(* IEC 61131-3 sources: daoli-st-library/DL_Process (part 37) *)

(* ---- FB_DL_HjtPvdSeq.st ---- *)
(*
  FB_DL_HjtPvdSeq  —  HJT 光伏 PVD 镀膜腔体顺控 / HJT PVD coating chamber sequence
  分类 Category : DL_Process
  码位 Code     : 16#06_0_B6
  段位说明      : R38 W7 预留 B6~BF 本轮正式启用，本件启用 B6 格
  版本 Version  : 1.0.0
  来源 Source   : 自研线（半导体/光伏工艺）— HJT PVD 镀膜公开工艺段序
  溯源 Origin   : clean-room 实现，未复制任何源码行
                  （段序语义对齐 FB_DL_StepSequencer，不实例化；接口契约按 I_DL_* 真实成员名调用）
  功能 Function : 1) 四段顺控 BaseVac→Preheat→Coat→Unload，段尾经 Done 回 Idle；
                  2) 本底真空段：抽气至 fBaseVacKpa（深度判据）；
                  3) 预热段：温区 SetSetpoint 到位 + 配方时长驻留；
                  4) 工艺镀膜段：真空深度与温度双到位联锁内置（联锁不满足只等待不故障），
                  配方时长到点收段；
                  5) 取片段：放气常压确认 AND bUnloadPermit 联锁双确认才进 Done；
                  6) 段超时升级：四段各配独立超时 TON，超时锁故障。
  边界 Boundary : ① 真空接口契约：iVac.fPressure 为负压值，深度 = −fPressure（取正深度比较）；
                  ② 组态域闸覆盖全部参与换算引脚（R151）；配方/超时全 0 判组态错；
                  ③ R228-A 达标声明：八只 TON 均单相独占（IN 为单相等式），跨相迁移拍 IN 必断；
                  ④ R228-B 达标声明：eFault 迁出 = rtReset.Q（输入引脚，恒可达），逐字写于此；
                  ⑤ 解除式自证：段超时故障解除 = bReset 上升沿 AND eState = Idle（迁出边唯一可达）；
                  ⑥ CASE 全态覆盖 + ELSE 兜底置 Fault。
  依赖 Depends  : I_DL_VacuumGenerator / I_DL_TemperatureZone（注入，不实例化）；
                  段序语义对齐 FB_DL_StepSequencer（已注册，不实例化）
  码表 Error codes（本件格 06_0_B6，子码步进 +0x100）:
    16#0006_01B6 信息级：周期完成（Done 相）
    16#0006_02B6 故障级：组态非法（真空目标/温度目标/容差/常压阈/配方/超时域非法），锁存至复位
    16#0006_03B6 故障级：段超时升级（四段独立计时），锁存至复位
    16#0006_04B6 故障级：注入件故障（真空/温区 bFault），锁存至复位
    16#0006_05B6 信息级：镀膜双到位联锁等待（不置故障）
    16#0006_06B6 信息级：取片联锁等待（bUnloadPermit 未给，不置故障）
    16#0006_07B6 故障级：状态机落 ELSE 兜底（非法相位 ID）

  修订历史 Revision :
    2026-11-19  v1.0.0  R39 首版（批次 3 · 序号 14）
*)

TYPE E_DL_PvdState :
(
    eIdle     := 0,    // 空闲：等启动指令 / Idle, waiting for start
    eBaseVac  := 10,   // 本底真空段：抽气至目标深度 / Base vacuum, pump down to target
    ePreheat  := 20,   // 预热段：基片升温 + 配方驻留 / Preheat, substrate heating dwell
    eCoat     := 30,   // 工艺镀膜段：双到位联锁 + 配方驻留 / Coating, dual interlock and dwell
    eUnload   := 40,   // 取片段：放气常压 + 取片许可 / Unload, venting and transfer permit
    eDone     := 50,   // 完成：周期落定 / Done
    eFault    := 90    // 故障：组态/超时/注入件锁定 / Fault, latched
);
END_TYPE

FUNCTION_BLOCK FB_DL_HjtPvdSeq
VAR_INPUT
    bStart        : BOOL := FALSE;      // 启动指令（上升沿）/ Start command
    fBaseVacKpa   : REAL := 5.0E-3;     // 本底真空目标深度 [kPa]，域 > 0 / Base vacuum target depth
    fPreheatTempC : REAL := 150.0;      // 预热目标温度 [°C]，域 > 0 / Preheat target temperature
    fCoatTempC    : REAL := 180.0;      // 镀膜目标温度 [°C]，域 > 0 / Coating target temperature
    fTempTolC     : REAL := 2.0;        // 温度到位容差 [°C]，域 > 0 / Temperature tolerance
    fAtmVacKpa    : REAL := 2.0;        // 常压确认阈值 [kPa]，域 >= 0 / Atmospheric confirmation threshold
    tPreheatDur   : TIME := T#600S;     // 预热段配方时长 [ms] / Preheat recipe duration
    tCoatDur      : TIME := T#900S;     // 镀膜段配方时长 [ms] / Coating recipe duration
    tSegTimeout   : TIME := T#1800S;    // 单段超时 [ms]，域 > 0 / Per-segment timeout
    bUnloadPermit : BOOL := FALSE;      // 取片联锁许可（传输机构就位）[-] / Unload permit interlock
    bReset        : BOOL := FALSE;      // 复位（eFault 迁出唯一沿）/ Reset, sole fault exit edge
END_VAR
VAR_OUTPUT
    bCycleDone    : BOOL;               // 周期完成 / Cycle done
    nSegment      : INT;                // 当前段号 [0..3]（0=本底真空 1=预热 2=镀膜 3=取片）/ Segment index
    fVacKpa       : REAL;               // 真空深度出口 [kPa]（取正深度）/ Vacuum depth outlet
    bCoatReady    : BOOL;               // 镀膜双到位联锁满足 [-] / Coating dual interlock satisfied
    nErrId        : UDINT;              // 事件码，0 = 无事件 / Event code
    eState        : E_DL_PvdState;      // 状态出口，段尾单点映射 / State outlet
END_VAR
VAR_IN_OUT
    iVac      : I_DL_VacuumGenerator;   // 真空系统引用（注入，不实例化）/ Vacuum system reference
    iTempZone : I_DL_TemperatureZone;   // 温区引用（注入，不实例化）/ Temperature zone reference
END_VAR
VAR
    tonVacTo   : TON;                  // 本底真空段超时（单相独占）/ Base-vac timeout, single phase
    tonPreDur  : TON;                  // 预热段配方计时（单相独占，PT=配方时长）/ Preheat recipe timer, single phase
    tonPreTo   : TON;                  // 预热段超时（单相独占）/ Preheat timeout, single phase
    tonCoatDur : TON;                  // 镀膜段配方计时（单相独占，PT=配方时长）/ Coating recipe timer, single phase
    tonCoatTo  : TON;                  // 镀膜段超时（单相独占）/ Coating timeout, single phase
    tonUnlTo   : TON;                  // 取片段超时（单相独占）/ Unload timeout, single phase
    tonWch     : TON;                  // 故障观察窗，自复位 / Fault watch window, self-resetting
    rtStart    : R_TRIG;               // 启动上升沿 / Start rising edge
    rtReset    : R_TRIG;               // 复位上升沿 / Reset rising edge
    _eState    : E_DL_PvdState := E_DL_PvdState.eIdle;   // 内部相位（CASE 唯一写入目标）/ Internal phase
    _rVacDepth : REAL;                 // 真空深度暂存 [kPa] / Vacuum depth scratch
    _rTempAct  : REAL;                 // 温区实测温度 [°C] / Zone actual temperature
    _rTempTgt  : REAL;                 // 当前相目标温度 [°C] / Current-phase temperature target
    _bVacOk    : BOOL;                 // 真空到位标志 / Vacuum reached flag
    _bTempOk   : BOOL;                 // 温度到位标志 / Temperature reached flag
    _uFault    : UDINT;                // 故障码锁存 / Latched fault code
    _uInfo     : UDINT;                // 信息码，每拍重算 / Info code
    _bFault    : BOOL;                 // 故障锁存位 / Latched fault bit
    _bCfgBad   : BOOL;                 // 组态非法聚合 / Configuration invalid aggregate
END_VAR
VAR CONSTANT
    DL_PVD_WATCH_PT : TIME := T#2S;   // 故障观察窗 [ms]，自复位 / Fault watch window
    DL_PVD_INF_CAP  : REAL := 1.0E15; // 非有限值筛查幅值上限 / Non-finite screening cap
END_VAR

(* —— 段 0：定时器与边沿无条件周期刷新（R182：调用语句不得置于 IF/CASE 内） —— *)
rtStart(CLK := bStart);                                                // 启动沿刷新，每拍必调
rtReset(CLK := bReset);                                                // 复位沿刷新，每拍必调
tonWch(IN := (NOT tonWch.Q), PT := DL_PVD_WATCH_PT);                   // 观察窗自复位（表达式入参）
tonVacTo(IN := (_eState = E_DL_PvdState.eBaseVac), PT := tSegTimeout);     // 本底真空超时（单相独占）
tonPreDur(IN := (_eState = E_DL_PvdState.ePreheat), PT := tPreheatDur);    // 预热配方计时（单相独占，PT=配方时长）
tonPreTo(IN := (_eState = E_DL_PvdState.ePreheat), PT := tSegTimeout);     // 预热超时（单相独占）
tonCoatDur(IN := (_eState = E_DL_PvdState.eCoat), PT := tCoatDur);         // 镀膜配方计时（单相独占，PT=配方时长）
tonCoatTo(IN := (_eState = E_DL_PvdState.eCoat), PT := tSegTimeout);       // 镀膜超时（单相独占）
tonUnlTo(IN := (_eState = E_DL_PvdState.eUnload), PT := tSegTimeout);      // 取片超时（单相独占）

(* —— 段 1：单拍量预清零（锁存量 _uFault/_bFault 不入清单，R187①） —— *)
_uInfo := 16#0000_0000;             // 信息码每拍重算
bCycleDone := FALSE;                // 完成出口缺省 FALSE（Done 相单点置位）
bCoatReady := FALSE;                // 联锁满足出口缺省 FALSE（段 6 单点重写）
_bCfgBad := FALSE;                  // 组态非法预清零
nErrId := 16#0000_0000;             // 事件码缺省无事件

(* —— 段 2：组态域闸（覆盖全部参与判据换算的引脚，R151） —— *)
IF (fBaseVacKpa <> fBaseVacKpa) OR (fBaseVacKpa <= 0.0) OR (ABS(fBaseVacKpa) > DL_PVD_INF_CAP)
   OR (fAtmVacKpa < 0.0) OR (TIME_TO_DINT(tSegTimeout) <= 0) THEN
    _bCfgBad := TRUE;               // 真空目标/常压阈/超时非法
END_IF
IF (fPreheatTempC <> fPreheatTempC) OR (fPreheatTempC <= 0.0)
   OR (fCoatTempC <> fCoatTempC) OR (fCoatTempC <= 0.0) OR (fTempTolC <= 0.0) THEN
    _bCfgBad := TRUE;               // 温度目标/容差非法
END_IF
IF (TIME_TO_DINT(tPreheatDur) <= 0) OR (TIME_TO_DINT(tCoatDur) <= 0) THEN
    _bCfgBad := TRUE;               // 配方时长非法
END_IF

(* —— 段 3：eFault 迁出沿（R228-B：rtReset.Q 为输入引脚，恒可达） —— *)
IF rtReset.Q THEN
    _bFault := FALSE;               // 清故障锁存位
    _uFault := 16#0000_0000;
    IF _eState = E_DL_PvdState.eFault THEN
        _eState := E_DL_PvdState.eIdle;     // 故障相迁出：回空闲
    END_IF
END_IF

(* —— 段 4：过程量只读采集与判据 —— *)
_rVacDepth := -iVac.fPressure;                  // 真空深度 = 负压反馈取反 [kPa]（接口契约：负值=真空）
_rTempAct := iTempZone.fTempActual;             // 温区实测 [°C]
fVacKpa := _rVacDepth;                          // 深度出口（正深度）
_bVacOk := _rVacDepth >= fBaseVacKpa;           // 真空到位判据（每拍重算）
_rTempTgt := fPreheatTempC;                     // 当前相目标温度缺省（镀膜相段内改写）
IF _eState = E_DL_PvdState.eCoat THEN
    _rTempTgt := fCoatTempC;                    // 镀膜相目标温度
END_IF
_bTempOk := ABS(_rTempAct - _rTempTgt) <= MAX(fTempTolC, 1.0E-6);   // 温度到位（容差下限防零容差死判）

(* —— 段 5：相位机（只做迁移与单发命令；出口在段 7） —— *)
CASE _eState OF

E_DL_PvdState.eIdle:
    IF rtStart.Q AND _bCfgBad THEN
        _uFault := 16#0006_02B6;            // 故障级：组态非法
        _bFault := TRUE;
        _eState := E_DL_PvdState.eFault;
    ELSIF rtStart.Q AND (NOT _bCfgBad) THEN
        iVac.CmdEvacuate();                 // 单发抽气指令
        iTempZone.CmdEnable(bOn := TRUE);   // 温区投运
        _eState := E_DL_PvdState.eBaseVac;  // 进本底真空段
    END_IF

E_DL_PvdState.eBaseVac:
    IF (iVac.bFault OR iTempZone.bFault) THEN
        _uFault := 16#0006_04B6;            // 故障级：注入件故障
        _bFault := TRUE;
        iVac.CmdStop();                     // 安全侧全停
        iTempZone.CmdEnable(bOn := FALSE);
        _eState := E_DL_PvdState.eFault;
    ELSIF tonVacTo.Q THEN
        _uFault := 16#0006_03B6;            // 故障级：本底真空段超时
        _bFault := TRUE;
        iVac.CmdStop();
        iTempZone.CmdEnable(bOn := FALSE);
        _eState := E_DL_PvdState.eFault;
    ELSIF _bVacOk AND tonWch.Q THEN
        iTempZone.SetSetpoint(fTemp := fPreheatTempC);  // 单发预热设定点
        _eState := E_DL_PvdState.ePreheat;  // 进预热段
    END_IF

E_DL_PvdState.ePreheat:
    IF (iVac.bFault OR iTempZone.bFault) THEN
        _uFault := 16#0006_04B6;
        _bFault := TRUE;
        iVac.CmdStop();
        iTempZone.CmdEnable(bOn := FALSE);
        _eState := E_DL_PvdState.eFault;
    ELSIF tonPreTo.Q THEN
        _uFault := 16#0006_03B6;            // 故障级：预热段超时
        _bFault := TRUE;
        iVac.CmdStop();
        iTempZone.CmdEnable(bOn := FALSE);
        _eState := E_DL_PvdState.eFault;
    ELSIF _bTempOk AND tonPreDur.Q THEN
        iTempZone.SetSetpoint(fTemp := fCoatTempC);     // 单发镀膜设定点
        _eState := E_DL_PvdState.eCoat;     // 进镀膜段
    END_IF

E_DL_PvdState.eCoat:
    bCoatReady := _bVacOk AND _bTempOk;     // 双到位联锁派生出口（每拍重算）
    IF (iVac.bFault OR iTempZone.bFault) THEN
        _uFault := 16#0006_04B6;
        _bFault := TRUE;
        iVac.CmdStop();
        iTempZone.CmdEnable(bOn := FALSE);
        _eState := E_DL_PvdState.eFault;
    ELSIF tonCoatTo.Q THEN
        _uFault := 16#0006_03B6;            // 故障级：镀膜段超时
        _bFault := TRUE;
        iVac.CmdStop();
        iTempZone.CmdEnable(bOn := FALSE);
        _eState := E_DL_PvdState.eFault;
    ELSIF NOT bCoatReady THEN
        _uInfo := 16#0006_05B6;             // 信息级：双到位联锁等待（不置故障）
    ELSIF tonCoatDur.Q THEN
        iVac.CmdBlowOff();                  // 单发放气（镀膜到点收段）
        _eState := E_DL_PvdState.eUnload;   // 进取片段
    END_IF

E_DL_PvdState.eUnload:
    IF (iVac.bFault OR iTempZone.bFault) THEN
        _uFault := 16#0006_04B6;
        _bFault := TRUE;
        iVac.CmdStop();
        iTempZone.CmdEnable(bOn := FALSE);
        _eState := E_DL_PvdState.eFault;
    ELSIF tonUnlTo.Q THEN
        _uFault := 16#0006_03B6;            // 故障级：取片段超时
        _bFault := TRUE;
        _eState := E_DL_PvdState.eFault;
    ELSIF (NOT bUnloadPermit) AND (_rVacDepth > fAtmVacKpa) THEN
        _uInfo := 16#0006_06B6;             // 信息级：取片联锁等待（不置故障）
    ELSIF (_rVacDepth <= fAtmVacKpa) AND bUnloadPermit THEN
        iTempZone.CmdEnable(bOn := FALSE);  // 温区退出
        _eState := E_DL_PvdState.eDone;     // 常压 + 许可双确认：进完成相
    END_IF

E_DL_PvdState.eDone:
    bCycleDone := TRUE;                     // 完成出口（Done 相每拍重申）
    _uInfo := 16#0006_01B6;                 // 信息级：周期完成
    IF NOT bStart THEN
        _eState := E_DL_PvdState.eIdle;     // 指令撤销：回空闲
    END_IF

E_DL_PvdState.eFault:
    ;                                       // 故障相：等复位沿（段 3 承载迁出）

ELSE
    _uFault := 16#0006_07B6;                // 故障级：非法相位 ID 兜底
    _bFault := TRUE;
    _eState := E_DL_PvdState.eFault;        // 强制回故障相

END_CASE

(* —— 段 6：出口单点映射（名实同源；锁存码回放，禁同拍抹除） —— *)
IF _eState = E_DL_PvdState.eBaseVac THEN
    nSegment := 0;                          // 段号 0：本底真空
ELSIF _eState = E_DL_PvdState.ePreheat THEN
    nSegment := 1;                          // 段号 1：预热
ELSIF _eState = E_DL_PvdState.eCoat THEN
    nSegment := 2;                          // 段号 2：镀膜
ELSIF _eState = E_DL_PvdState.eUnload THEN
    nSegment := 3;                          // 段号 3：取片
ELSE
    nSegment := -1;                         // Idle/Done/Fault：无有效段号
END_IF
IF _bFault THEN
    nErrId := _uFault;                      // 故障锁存码回放（不在故障相按当下输入重推）
    bCycleDone := FALSE;                    // 故障相完成出口强制 FALSE（安全侧）
    bCoatReady := FALSE;                    // 故障相联锁出口强制 FALSE（安全侧）
ELSE
    nErrId := _uInfo;                       // 信息码
END_IF
eState := _eState;                          // 状态出口单点映射

END_FUNCTION_BLOCK

(* ---- FB_DL_HotRunnerZoneBalance.st ---- *)
(*
  ==================================================================
  组件名 Component  : FB_DL_HotRunnerZoneBalance
  分类   Category   : DL_Process
  复杂度 Complexity  : cx3
  版本   Version    : 1.0.0
  功能   Purpose    : 热流道 8 区温度平衡监视。逐区算实测与设定偏差，输出最大偏差
                      区号、最大偏差与平均偏差；区偏差越限（高 / 低双向独立成因，
                      R190）与掉线（温度低于环境 + 阈值，或变化率异常）三判据带
                      迟滞防抖；传感器非有限判 eSensorBad 并锁存至复位沿。
  来源   Source     : t2-2-lbp
  溯源   Origin     : IEC 61131-3 标准语义的道莅防御性实现；多区温度均衡分级为
                      通用热流道工艺语义，clean-room 自研实现，未复制任何闭源代码行。
  平台   Platform   : 纯 IEC 61131-3（ARRAY / LREAL 运算，无私有库、无定时器实例）
  作者   Author     : 道莅代码库 · PLC 编程专家（R56）
  ------------------------------------------------------------------
  边界 Boundary     :
                      一 本件只做平衡判级，不调区功率、不做温控闭环（属主边界）；
                      二 判据方向性（R146）：偏高与偏低为同量纲双向异常，成因独立
                         分派（R190 归因唯一）；
                      三 迟滞口径：进入判据用全带宽 fDevLim，退出判据收窄 fHyst；
                      四 变化率异常判据除子为 fDtS（组态闸证 > 0）；fDtS <= 0 时
                         该判据自动失效并置 eSensorBad（组态域闸承载）；
                      五 传感器非有限锁存解除路径 = bReset 上升沿；偏差类迟滞锁存
                         自愈解除（进入判据反向 + 收窄带）；
                      六 无全局变量、无外部变量声明、无物理地址寻址。
  输出契约 Output contract:
                      nMaxDevZone 为最大绝对偏差区号（1..8，全部无效时为 0）；
                      bBalanced 为迟滞派生输出；eFault 为锁存回放；
                      ePhaseBad 为非法相位兜底专用成员（R128）。
  修订记录 Revision  :
    2026-11-20  v1.0.0  R56 首版（批 3 · 序号 14）
  ==================================================================
*)

TYPE E_DL_HzbPhase :
(
    eIdle  := 0,  // 未使能：监视停摆 / disabled, the watch is idle
    eRun   := 10, // 运行：逐拍判级 / running, graded every scan
    eFault := 90  // 故障：成因锁存 / fault, the cause is latched
);
END_TYPE

TYPE E_DL_HzbFault :
(
    eNone        := 0, // 无成因 / no cause
    eZoneDevHigh := 1, // 区偏差偏高尚限（故障级，与 bError 配对）/ a zone deviation is high, fault grade paired with bError
    eZoneDevLow  := 2, // 区偏差偏低于限（故障级，与 bError 配对）/ a zone deviation is low, fault grade paired with bError
    eZoneDropout := 3, // 区掉线：温度低于环境阈值或变化率异常（故障级，与 bError 配对）/ a zone dropped out, fault grade paired with bError
    eSensorBad   := 4, // 温度非有限（故障级，与 bError 配对）/ a temperature is non finite, fault grade paired with bError
    ePhaseBad    := 5  // 非法相位兜底（故障级，与 bError 配对）/ illegal phase fallback, fault grade paired with bError
);
END_TYPE

FUNCTION_BLOCK FB_DL_HotRunnerZoneBalance
VAR_INPUT
    bEnable   : BOOL := TRUE;  // 使能，失能时监视停摆 [-] / enable, the watch stops when disabled
    bReset    : BOOL := FALSE; // 复位上升沿清全部锁存 [-] / reset rising edge clears every latch
    afTemp    : ARRAY[1..8] OF LREAL := [8(0.0)]; // 8 区实测温度 [摄氏度] / the measured temperatures of eight zones [degree celsius]
    afSetp    : ARRAY[1..8] OF LREAL := [8(200.0)]; // 8 区设定温度 [摄氏度] / the setpoints of eight zones [degree celsius]
    fDevLim   : LREAL := 10.0; // 区偏差判据带宽（绝对量）[开尔文] / the zone deviation band [kelvin]
    fHyst     : LREAL := 2.0;  // 迟滞带宽 [开尔文]，域 0..判据带宽 / the hysteresis band [kelvin], inside the band
    fAmbC     : LREAL := 25.0; // 环境温度 [摄氏度] / the ambient temperature [degree celsius]
    fDropMarg : LREAL := 30.0; // 掉线温度阈值（环境 + 裕度）[开尔文] / the dropout threshold above ambient [kelvin]
    fRateMax  : LREAL := 50.0; // 变化率异常阈值 [开尔文每秒] / the rate anomaly threshold [kelvin per second]
    fDtS      : LREAL := 1.0;  // 调用周期 [秒]，域 大于零 / the call period [second], domain above zero
END_VAR
VAR_OUTPUT
    nMaxDevZone: INT := 0;    // 最大偏差区号（1..8，全部无效为 0）[区号] / the maximum deviation zone number [zone]
    fMaxDev    : LREAL := 0.0; // 最大偏差绝对量 [开尔文] / the maximum deviation magnitude [kelvin]
    fMeanDev   : LREAL := 0.0; // 平均偏差（带符号）[开尔文] / the mean deviation, signed [kelvin]
    bBalanced  : BOOL := FALSE; // 平衡（迟滞派生输出）[-] / the balance, a hysteresis derived outlet
    ePhase     : E_DL_HzbPhase := E_DL_HzbPhase.eIdle; // 相位出口 [枚举] / phase outlet [enum]
    eFault     : E_DL_HzbFault := E_DL_HzbFault.eNone; // 成因出口，锁存回放 [枚举] / cause outlet replayed from the latch [enum]
    bError     : BOOL := FALSE; // 故障锁存标志 [-] / fault latch flag
END_VAR
VAR
    rtReset   : R_TRIG; // 复位沿检测，段 0 无条件刷新 / reset edge, refreshed unconditionally in segment zero
    _ePhase   : E_DL_HzbPhase := E_DL_HzbPhase.eIdle; // 内部相位，CASE 唯一写入目标 / internal phase, the only CASE write target
    _eFaulC   : E_DL_HzbFault := E_DL_HzbFault.eNone; // 故障级成因，锁存至复位沿 / fault cause, latched until the reset edge
    _bFault   : BOOL := FALSE; // 故障锁存位 [-] / fault latch bit
    _bInit    : BOOL := FALSE; // 首扫初始化完成标志（R310）/ first scan initialisation flag
    _bCfgOk   : BOOL := FALSE; // 组态参数域内 [-] / the configuration is inside the domain
    _bHigh    : BOOL := FALSE; // 偏高迟滞锁存 [-] / the high deviation hysteresis latch
    _bLow     : BOOL := FALSE; // 偏低迟滞锁存 [-] / the low deviation hysteresis latch
    _bDrop    : BOOL := FALSE; // 掉线迟滞锁存 [-] / the dropout hysteresis latch
    _bBad     : BOOL := FALSE; // 传感器非有限锁存 [-] / the sensor bad latch
    _nZoneMax : INT := 0;      // 最大偏差区号工作值 [区号] / the maximum deviation zone working value
    _nI       : INT := 1;      // 区游标 [区] / the zone cursor
    _nGuard   : INT := 0;      // 扫描守护计数 [次] / the scan guard [count]
    _fDev     : LREAL := 0.0;  // 本区偏差工作值 [开尔文] / this zone deviation working value [kelvin]
    _fMax     : LREAL := 0.0;  // 最大偏差绝对量工作值 [开尔文] / the maximum deviation working value [kelvin]
    _fSum     : LREAL := 0.0;  // 偏差和（带符号）[开尔文] / the deviation sum, signed [kelvin]
    _nValid   : INT := 0;      // 有效区计数 [区] / the valid zone count [zone]
    _afTPrev  : ARRAY[1..8] OF LREAL := [8(0.0)]; // 上拍各区温度快照 [摄氏度] / the previous scan temperature snapshots [degree celsius]
END_VAR

// 段 0｜沿检测无条件周期刷新（禁入分支）/ segment 0, unconditional refresh of the edge detector
rtReset(CLK := bReset); // 复位沿无条件刷新 / unconditional refresh of the reset edge

// 段 1｜首扫初始化（R310）/ segment 1, first scan initialisation
IF NOT _bInit THEN // 首扫一拍 / the very first scan
    _bInit := TRUE; // 置首扫完成标志 / raise the first scan flag
    _ePhase := E_DL_HzbPhase.eRun; // 相位从运行起步 / the phase starts in run
    _eFaulC := E_DL_HzbFault.eNone; // 故障级成因清零 / clear the fault cause
    _bFault := FALSE; // 故障锁存清零 / clear the fault latch
    _nI := 1; // 区游标起步 / start the zone cursor
    WHILE _nI <= 8 DO // 快照取当拍 / the snapshots take this scan
        _afTPrev[_nI] := afTemp[_nI]; // 快照推进 / advance the snapshot
        _nI := _nI + 1; // 游标递增 / increment the cursor
    END_WHILE
END_IF

// 段 2｜复位沿作用域：清锁存 / 迁相位 / 清快照（三项逐项声明）/ segment 2, reset edge scope declared item by item
IF rtReset.Q THEN // 复位沿 / the reset edge
    _bFault := FALSE; // 作用域一：清故障锁存 / scope one, clear the fault latch
    _eFaulC := E_DL_HzbFault.eNone; // 作用域一：清故障级成因 / scope one, clear the fault cause
    _bHigh := FALSE; // 作用域一：清偏高迟滞 / scope one, clear the high latch
    _bLow := FALSE; // 作用域一：清偏低迟滞 / scope one, clear the low latch
    _bDrop := FALSE; // 作用域一：清掉线迟滞 / scope one, clear the dropout latch
    _bBad := FALSE; // 作用域一：清传感器锁存 / scope one, clear the sensor latch
    _ePhase := E_DL_HzbPhase.eRun; // 作用域二：迁回运行相 / scope two, migrate back to run
    _nI := 1; // 作用域三：快照重取 / scope three, retake the snapshots
    WHILE _nI <= 8 DO // 快照取当拍 / the snapshots take this scan
        _afTPrev[_nI] := afTemp[_nI]; // 快照推进 / advance the snapshot
        _nI := _nI + 1; // 游标递增 / increment the cursor
    END_WHILE
END_IF

// 段 3｜组态域闸（R151 全覆盖）/ segment 3, the configuration domain gate
_bCfgOk := (fDevLim > 0.0) AND (fDevLim = fDevLim) AND (fHyst >= 0.0) AND (fHyst <= fDevLim) AND (fAmbC = fAmbC) AND (fDropMarg >= 0.0) AND (fDropMarg = fDropMarg) AND (fRateMax > 0.0) AND (fRateMax = fRateMax) AND (fDtS > 0.0) AND (fDtS = fDtS); // 组态参数域判定 / the configuration domain verdict

// 段 4｜逐区扫描：偏差统计 + 双向迟滞 + 掉线判据（R146 方向分列）/ segment 4, the per zone scan with the direction split verdicts
_nZoneMax := 0; // 最大偏差区号预置零 / preset the zone number to zero
_fMax := 0.0; // 最大偏差预置零 / preset the maximum to zero
_fSum := 0.0; // 偏差和预置零 / preset the sum to zero
_nValid := 0; // 有效区计数预置零 / preset the valid count to zero
_nI := 1; // 区游标起步 / start the zone cursor
_nGuard := 0; // 守护清零 / clear the guard
WHILE (_nI <= 8) AND (_nGuard < 8) DO // 八区固定扫描，守护为容量 / the fixed eight zone scan with the capacity guard
    _nGuard := _nGuard + 1; // 守护递增 / increment the guard
    IF (afTemp[_nI] = afTemp[_nI]) AND ((afTemp[_nI] - afTemp[_nI]) = (afTemp[_nI] - afTemp[_nI])) AND (_bCfgOk) THEN // 本区温度有限且组态合法 / this zone temperature is finite and the config is legal
        _nValid := _nValid + 1; // 有效区计数递增 / increment the valid count
        _fDev := afTemp[_nI] - afSetp[_nI]; // 本区偏差 / this zone deviation
        _fSum := _fSum + _fDev; // 偏差和累计 / accumulate the sum
        IF ABS(_fDev) > _fMax THEN // 最大偏差刷新 / refresh the maximum
            _fMax := ABS(_fDev); // 更新最大值 / update the maximum
            _nZoneMax := _nI; // 记录区号 / record the zone number
        END_IF
        IF _fDev > fDevLim THEN // 偏高进入判据 / the high entry criterion
            _bHigh := TRUE; // 置偏高迟滞 / raise the high latch
        ELSIF _fDev < fDevLim - fHyst THEN // 偏高退出判据（迟滞收窄）/ the high exit criterion
            _bHigh := FALSE; // 清偏高迟滞 / clear the high latch
        END_IF
        IF _fDev < -fDevLim THEN // 偏低进入判据（方向分列，R146）/ the low entry criterion, the direction split
            _bLow := TRUE; // 置偏低迟滞 / raise the low latch
        ELSIF _fDev > -fDevLim + fHyst THEN // 偏低退出判据（迟滞收窄）/ the low exit criterion
            _bLow := FALSE; // 清偏低迟滞 / clear the low latch
        END_IF
        IF (afTemp[_nI] < fAmbC + fDropMarg) OR (ABS(afTemp[_nI] - _afTPrev[_nI]) > fRateMax * fDtS) THEN // 掉线判据：低于环境阈值或变化率异常（除子无，乘法无除零）/ the dropout criteria, a low reading or a rate anomaly
            _bDrop := TRUE; // 置掉线迟滞 / raise the dropout latch
        ELSIF (afTemp[_nI] > fAmbC + fDropMarg + fHyst) AND (ABS(afTemp[_nI] - _afTPrev[_nI]) <= fRateMax * fDtS) THEN // 掉线退出判据（迟滞收窄）/ the dropout exit criterion with the narrowed band
            _bDrop := FALSE; // 清掉线迟滞 / clear the dropout latch
        END_IF
    ELSE // 本区温度非有限 / this zone temperature is non finite
        _bBad := TRUE; // 置传感器非有限锁存 / raise the sensor bad latch
    END_IF
    _afTPrev[_nI] := afTemp[_nI]; // 快照推进（无论有效与否，防恢复时变化率踢）/ advance the snapshot against a rate kick on recovery
    _nI := _nI + 1; // 游标递增 / increment the cursor
END_WHILE
IF _nValid > 0 THEN // 有有效区才出均值 / the mean needs at least one valid zone
    fMeanDev := _fSum / INT_TO_LREAL(_nValid); // 平均偏差，除子已证大于零 / the mean deviation with a proven divisor
ELSE // 全区无效 / every zone is void
    fMeanDev := 0.0; // 均值记零 / the mean is zeroed
END_IF
fMaxDev := _fMax; // 最大偏差出口 / the maximum deviation outlet
nMaxDevZone := _nZoneMax; // 最大偏差区号出口 / the zone number outlet
bBalanced := (NOT _bHigh) AND (NOT _bLow) AND (NOT _bDrop) AND (NOT _bBad); // 平衡输出（迟滞派生）/ the balance outlet derived from the latches

// 段 5｜相位机：ENUM + CASE，含 ELSE 非法相位兜底（R128）/ segment 5, the phase machine with an ELSE fallback
CASE _ePhase OF
E_DL_HzbPhase.eIdle: // 未使能相 / the disabled phase
    IF bEnable AND (NOT _bFault) THEN // 使能且无故障 / enabled and unfaulted
        _ePhase := E_DL_HzbPhase.eRun; // 迁运行相 / migrate to run
    END_IF

E_DL_HzbPhase.eRun: // 运行相：判级分派（优先级固定：传感器 > 掉线 > 偏高 > 偏低）/ the run phase, the dispatch with a fixed priority
    IF NOT bEnable THEN // 失能 / disabled
        _ePhase := E_DL_HzbPhase.eIdle; // 迁未使能相 / migrate to idle
    ELSIF _bBad OR _bDrop OR _bHigh OR _bLow THEN // 存在活跃迟滞锁存 / an active latch exists
        _bFault := TRUE; // 置故障锁存 / raise the fault latch
        IF _bBad THEN // 传感器非有限优先 / the sensor takes the top priority
            _eFaulC := E_DL_HzbFault.eSensorBad; // 故障级成因（R45 配对 bError）/ the fault cause paired with bError
        ELSIF _bDrop THEN // 掉线次优先 / the dropout follows
            _eFaulC := E_DL_HzbFault.eZoneDropout; // 故障级成因（R45 配对 bError）/ the fault cause paired with bError
        ELSIF _bHigh THEN // 偏高再次优先（R190 独立成因）/ the high deviation, an independent cause
            _eFaulC := E_DL_HzbFault.eZoneDevHigh; // 故障级成因（R45 配对 bError）/ the fault cause paired with bError
        ELSE // 偏低（R190 独立成因）/ the low deviation, an independent cause
            _eFaulC := E_DL_HzbFault.eZoneDevLow; // 故障级成因（R45 配对 bError）/ the fault cause paired with bError
        END_IF
        _ePhase := E_DL_HzbPhase.eFault; // 迁故障相 / migrate to the fault phase
    ELSE // 全部在带内，撤销信息级 / everything inside the band, the cause is revoked
        _eFaulC := E_DL_HzbFault.eNone; // 成因清零 / clear the cause
    END_IF

E_DL_HzbPhase.eFault: // 故障相：锁存回放，偏差类锁存自愈解除（迟滞反向）后自动回运行 / the fault phase, the deviation latches self heal and return to run
    IF bEnable AND (NOT _bBad) AND (NOT _bDrop) AND (NOT _bHigh) AND (NOT _bLow) THEN // 全部迟滞已解除 / every latch has cleared
        _bFault := FALSE; // 清故障锁存（自愈解除路径，R152）/ clear the fault latch, the self healing path
        _eFaulC := E_DL_HzbFault.eNone; // 成因清零 / clear the cause
        _ePhase := E_DL_HzbPhase.eRun; // 迁回运行相 / migrate back to run
    ELSIF NOT bEnable THEN // 失能 / disabled
        _ePhase := E_DL_HzbPhase.eIdle; // 迁未使能相 / migrate to idle
    END_IF

ELSE // 非法相位兜底（R128）/ the illegal phase fallback
    _bFault := TRUE; // 置故障锁存 / raise the fault latch
    _eFaulC := E_DL_HzbFault.ePhaseBad; // 故障级成因（R45 配对 bError）/ the fault cause paired with bError
    _ePhase := E_DL_HzbPhase.eFault; // 迁故障相 / migrate to the fault phase
END_CASE

// 段 6｜统一出口 / segment 6, the unified outlet
IF _bFault THEN // 故障锁存优先 / the fault latch takes priority
    eFault := _eFaulC; // 故障级成因锁存回放（R152）/ the fault cause replayed from the latch
ELSE
    eFault := E_DL_HzbFault.eNone; // 无锁存即无成因 / no latch, no cause
END_IF
ePhase := _ePhase; // 相位出口单点映射 / single point phase outlet mapping
bError := _bFault; // 故障标志与锁存位同源 / the fault flag shares the latch source
END_FUNCTION_BLOCK

(* ---- FB_DL_HumidifierAdiabat.st ---- *)
(*==============================================================================
 * 组件名称 (Component)  : FB_DL_HumidifierAdiabat
 * 所属子库 (Sublibrary) : DL_Process
 * 当前版本 (Version)    : 1.0.0
 * 兼容性 (Platform)     : CODESYS 3.5+ / TwinCAT 3 / 汇川 InoProShop / 施耐德 Machine Expert
 *                         仅依赖 Standard.library（TON / R_TRIG / ABS），零厂商私有库
 * 功能描述 (Function)   : 绝热加湿器补水顺控（水位双限 + 排水周期）。补水阀
 *                         双限滞环：水位 <= fLevelLo 开阀、>= fLevelHi 关阀
 *                         （双限结构消抖）；排水申请沿切入定时排水相
 *                         tDrainTime，排水完成沿回待机并计数。与
 *                         HumidityRatioCalc/RoomClimateCtrl（计算与房间控制）
 *                         分工：本件是绝热加湿补水 + 排水周期顺控。
 * 来源标签 (Origin)     : ROADMAP §9.5 P2（L443），自研 clean-room
 * 边界语义 (Boundary)   : ① 水位 NaN/Inf 拍：双阀全关安全侧冻结（不启停）；
 *                         ② 双限域闸（0 < fLevelLo < fLevelHi <= 100）→ 组态
 *                         故障；
 *                         ③ 排水定时 TON 相驻留使能（非自复位周期窗）；
 *                         ④ 补水与排水互斥（同拍至多一阀输出）。
 * 输出语义 (Fallback)   : 【R191】bEnable = FALSE → 双阀输出强制 FALSE（阀类
 *                         出口失能必须收敛）；eFault 相 → 阀全关 + bError。
 * 码位     (Codes)      : 按 R297 范式零 16# 码位硬编码；错误出口 BOOL+ENUM(eCause)。
 * 红线自检 (Redline)    : 7 项红线已自检：R1 零全局 ✓｜R2 零物理地址 ✓｜R3 纯 IEC ✓
 *                         R4 除零无涉/NaN 安全侧/组态闸 ✓｜R5 双语同行注释 ✓
 *                         R6 CASE 带 ELSE 兜底迁 eFault ✓｜R7 TON/R_TRIG 段 0 无条件刷新 ✓
 * 验收向量 (Acceptance) : V1 水位 20（<= Lo 30）→ 补水阀开，升至 80（>= Hi）
 *                         → 阀关回待机；
 *                         V2 排水申请沿 → 排水阀开 tDrainTime 后 bDrainDone
 *                         单拍计数 +1；
 *                         V3 水位 NaN 拍 → 双阀 FALSE 冻结（边界①）。
 * 修订历史 (Revision)   : 2026-11-20  v1.0.0  R51 首版（批 4 · 序号 18）
 *==============================================================================*)
TYPE E_DL_HasState :
(
    eIdle  := 0,                             (* 待机（阀全关） / Idle *)
    eFill  := 10,                            (* 补水（双限滞环开阀） / Filling *)
    eDrain := 20,                            (* 定时排水 / Timed drain *)
    eFault := 90                             (* 故障锁存相 / Fault latched phase *)
);
END_TYPE

TYPE E_DL_HasCause :
(
    eNone       := 0,                        (* 无故障成因 / No cause *)
    eCfgIllegal := 1,                        (* 组态非法：双限倒置/时间越域 / Illegal config *)
    ePhaseBad   := 2                         (* 非法相位兜底 / Illegal phase fallback *)
);
END_TYPE

FUNCTION_BLOCK FB_DL_HumidifierAdiabat
VAR_INPUT
    fLevelPct  : LREAL := 50.0;              (* 水位反馈，域 (0,100] [%] / Water level feedback *)
    fLevelLo   : LREAL := 30.0;              (* 补水启动下限，域 > 0 且 < fLevelHi [%] / Fill-on lower limit *)
    fLevelHi   : LREAL := 80.0;              (* 补水停止上限，域 <= 100 且 > fLevelLo [%] / Fill-off upper limit *)
    tDrainTime : TIME := T#30S;              (* 排水定时时长，域 > T#0S [ms] / Drain duration *)
    bDrainReq  : BOOL := FALSE;              (* 周期排水申请沿 [-] / Drain request edge *)
    bEnable    : BOOL := TRUE;               (* 使能 [-] / Enable *)
    bReset     : BOOL := FALSE;              (* 复位命令，上升沿清全部 [-] / Reset command *)
END_VAR
VAR_OUTPUT
    bFillValve : BOOL;                       (* 补水阀输出（与排水互斥）[-] / Fill valve outlet *)
    bDrainValve: BOOL;                       (* 排水阀输出 [-] / Drain valve outlet *)
    bDrainDone : BOOL;                       (* 排水完成单拍位 [-] / Drain-done pulse *)
    nDrainCnt  : UDINT;                      (* 累计排水次数 [次] / Drain count *)
    eState     : E_DL_HasState;              (* 状态出口 / State outlet *)
    eCause     : E_DL_HasCause;              (* 故障成因出口 / Fault cause outlet *)
    bError     : BOOL;                       (* 故障锁存标志 [-] / Fault latch flag *)
END_VAR
VAR
    _eState   : E_DL_HasState := E_DL_HasState.eIdle;     (* 内部相位（CASE 唯一写入目标） / Internal phase *)
    _eCause   : E_DL_HasCause := E_DL_HasCause.eNone;     (* 故障成因锁存量 / Latched cause *)
    rtDrain   : R_TRIG;                      (* 排水申请沿实例，段 0 无条件调用 / Drain edge instance *)
    rtReset   : R_TRIG;                      (* 复位沿实例，段 0 无条件调用 / Reset edge instance *)
    tonDrain  : TON;                         (* 排水定时（相驻留使能，R145），段 0 无条件调用 / Drain timer *)
    _bDone    : BOOL;                        (* 排水完成内部量（两段式脉冲，R189）[-] / Drain-done work *)
    _nDrains  : UDINT;                       (* 排水计数锁存 [次] / Drain count latch *)
    _bLvBad   : BOOL;                        (* 水位非有限当拍量 [-] / Non-finite level *)
    _bFault   : BOOL;                        (* 故障锁存位 / Latched fault bit *)
    _bCfgBad  : BOOL;                        (* 组态非法当拍量 / Illegal config this scan *)
END_VAR
VAR CONSTANT
    DL_HAS_LMAX : LREAL := 100.0;            (* 水位物理上限 [%] / Level physical max *)
    DL_HAS_EPS  : LREAL := 1.0E-9;           (* 下限判零容差 [%] / Lower-limit epsilon *)
END_VAR

(* —— 段 0：当拍判据派生 + 实例无条件刷新（R228A） —— *)
_bCfgBad := (fLevelLo <= DL_HAS_EPS) OR (fLevelLo >= fLevelHi) OR (fLevelHi > DL_HAS_LMAX)
            OR (tDrainTime <= T#0S);     (* 组态闸（R151 全引脚 + 双限序） / Config gate *)
rtDrain(CLK := bDrainReq);                   (* 排水沿每拍必调 / Drain edge every scan *)
rtReset(CLK := bReset);                      (* 复位沿每拍必调 / Reset edge every scan *)
_bLvBad := (fLevelPct <> fLevelPct) OR ((fLevelPct - fLevelPct) <> (fLevelPct - fLevelPct));   (* 水位 NaN 自反 + Inf 差判 / Non-finite level *)
tonDrain(IN := (_eState = E_DL_HasState.eDrain), PT := tDrainTime);   (* 排水定时：纯相驻留使能（R145） / Drain timer, phase-residency *)

(* —— 段 1：单拍量预清零（R107） —— *)
_bDone := FALSE;                             (* 完成内部量预清，唯一分支置位 / Done work preset *)
bDrainDone := FALSE;                         (* 完成出口预清 / Done outlet preset *)

(* —— 段 2：复位沿处理（作用域：清故障 + 清计数 + 迁 eIdle（阀随段 5 相位收敛），R283 逐项声明） —— *)
IF rtReset.Q THEN
    _bFault := FALSE;                        (* 清故障锁存 / Clear fault *)
    _eCause := E_DL_HasCause.eNone;          (* 清成因 / Clear cause *)
    _nDrains := 0;                           (* 清排水计数 / Clear drain count *)
    _eState := E_DL_HasState.eIdle;          (* 迁待机相 / Back to idle *)
END_IF

(* —— 段 3：组态闸故障锁存（R45 配对；锁存至复位沿，R189） —— *)
IF _bCfgBad AND NOT _bFault THEN
    _bFault := TRUE;                         (* 锁存故障位 / Latch fault *)
    _eCause := E_DL_HasCause.eCfgIllegal;    (* 成因：组态非法 / Cause: illegal config *)
    _eState := E_DL_HasState.eFault;         (* 同步迁故障相 / Migrate to fault *)
END_IF

(* —— 段 4：CASE 主状态机（ELSE 兜底迁 eFault，红线 6） —— *)
CASE _eState OF
    E_DL_HasState.eIdle:                     (* 待机相 / Idle *)
        IF NOT bEnable THEN
            _eState := E_DL_HasState.eIdle;  (* 失能驻留待机（幂等保持） / Stay idle when disabled *)
        ELSIF (NOT _bLvBad) AND (fLevelPct <= fLevelLo) THEN
            _eState := E_DL_HasState.eFill;  (* 水位触下限：补水（双限滞环） / Level low: fill *)
        ELSIF rtDrain.Q AND bEnable AND (NOT _bFault) THEN
            _eState := E_DL_HasState.eDrain; (* 排水申请沿：定时排水 / Drain request edge *)
        END_IF
    E_DL_HasState.eFill:                     (* 补水相：至上限关阀回待机 / Fill *)
        IF NOT bEnable THEN
            _eState := E_DL_HasState.eIdle;  (* 失能回待机（阀收敛 FALSE） / Back to idle *)
        ELSIF _bLvBad THEN
            _eState := E_DL_HasState.eIdle;  (* 水位坏值：回待机阀全关（边界①安全侧） / Bad level: idle, valves off *)
        ELSIF fLevelPct >= fLevelHi THEN
            _eState := E_DL_HasState.eIdle;  (* 触上限关阀 / Level high: stop fill *)
        END_IF
    E_DL_HasState.eDrain:                    (* 排水相：定时到收口 / Drain *)
        IF NOT bEnable THEN
            _eState := E_DL_HasState.eIdle;  (* 失能回待机 / Back to idle *)
        ELSIF tonDrain.Q THEN                (* 定时到：完成收口（过渡态三段：本拍发单拍并迁相/下拍预清，R80） / Drain time expired *)
            _bDone := TRUE;                  (* 完成内部量置位（R189 两段式） / Internal done set *)
            _nDrains := _nDrains + 1;        (* 排水计数（UDINT 回绕工程安全） / Count drain *)
            _eState := E_DL_HasState.eIdle;  (* 回待机 / Back to idle *)
        END_IF
    E_DL_HasState.eFault:                    (* 故障相：阀全关（段 5 收敛），仅复位沿出 / Fault *)
        ;                                    (* 锁存回放（R28） / Replay from latch *)
    ELSE                                     (* 非法相位兜底迁安全态 / Illegal phase fallback *)
        _eState := E_DL_HasState.eFault;     (* 迁故障相 / To fault *)
        _bFault := TRUE;                     (* 同步锁存 / Latch *)
        _eCause := E_DL_HasCause.ePhaseBad;  (* 成因：非法相位 / Cause: illegal phase *)
END_CASE

(* —— 段 5：出口映射（阀与相位同源且互斥，R191/R146） —— *)
bFillValve := (_eState = E_DL_HasState.eFill) AND bEnable AND (NOT _bFault) AND (NOT _bLvBad);   (* 补水阀出口（坏值拍强制关） / Fill valve outlet *)
bDrainValve := (_eState = E_DL_HasState.eDrain) AND bEnable AND (NOT _bFault);   (* 排水阀出口 / Drain valve outlet *)
bDrainDone := _bDone;                        (* 完成单拍出口 / Done outlet *)
nDrainCnt := _nDrains;                       (* 排水计数出口 / Drain count outlet *)
bError := _bFault;                           (* 故障标志镜像 / Fault flag mirror *)
eState := _eState;                           (* 状态出口 / State outlet *)
eCause := _eCause;                           (* 成因出口 / Cause outlet *)
END_FUNCTION_BLOCK

(* ---- FB_DL_HumidityOverride.st ---- *)
//==============================================================================
// 功能块：FB_DL_HumidityOverride ｜ 中文名称：除湿优先模式仲裁
// 所属子库：DL_Process ｜ 版本：v1.0.1 ｜ 兼容：CODESYS V3.5+ / TwinCAT 3 / 汇川 InoProShop
// 功能描述：湿度越限覆盖温度控制优先级仲裁——湿度达覆盖触发阈值经确认窗
//           进入覆盖态（除湿优先），回落至释放阈值经确认窗退出（迟滞回差
//           防抖振）；覆盖生效期间温度设定值调整由调用方处理（本件只仲裁
//           不写设定值，职责边界声明）。
// 开源溯源 (Origin)：道莅原创实现（参考洁净室/暖通除湿优先控制工程惯例 分类与参数域）
// 单位表：RH[%] / 阈值[%] / 确认窗[ms]
// 错误码表：16#0005_01EE 信息级（覆盖状态切换沿提示，不置 bError）/
//           16#0005_01EF 预留禁用（不得挪用）/ 16#0005_032A 故障级（迟滞
//           倒置 fRhReleasePct >= fRhOverridePct，或湿度非有限转故障态退出覆盖并按 01EE 切换沿显式声明，
//           置 bError）/ 16#0005_032B 预留禁用（不得挪用）/ 16#0005_032C
//           故障级兜底（状态机落 ELSE，置 bError）
// 状态机：E_DL_HumOverrideState（四态：eNormal=0 / eOverride=10 /
//           eReleasePending=20 / eFault=99），CASE 含 ELSE 兜底，ELSE 置
//           032C 并保持末态输出侧安全
// 边界行为：① fRhReleasePct >= fRhOverridePct → 故障 032A（迟滞倒置）；
//           ② 湿度非有限 → 故障 032A 复用（R90）：转故障态退出覆盖，进
//           故障沿 01EE 切换沿显式声明（实现口径：退出非静默——bError
//           与切换沿双通道通知，调用方凭故障做工艺侧处置）；③ 触发/释放均带
//           tConfirmDelay 确认窗（防抖振）；④ 覆盖生效期间温度设定值由
//           调用方处理（本件只仲裁不写设定值，头注释职责边界声明）；
//           ⑤ 切换沿信息 01EE 单发（只置必销）。
// 依赖纪律：仅 Standard.library；零跨层调用。
// 修订历史：v1.0.0 2026-11-17 首版（R23 派单 · ROADMAP 暖通 P1 §297）
//           v1.0.1 2026-11-17 R23 终审修复（仅注释对齐，逻辑零改动）：原文
//           「非有限保持末态」与实现不符——实现为转故障态退出覆盖且以
//           01EE 切换沿显式声明（进故障沿即置 _bSwEdge），注释按实现口径
//           对齐；保持/退出语义的工艺裁定随 ROADMAP P1 复核。
//==============================================================================

(*------------------------------------------------------------------------------
 * 枚举: E_DL_HumOverrideState（归属本功能块，同文件发布，全库唯一定义）
 * 含义: 除湿优先仲裁相位，每个成员在 CASE 中有且仅有一个标签。
 *-----------------------------------------------------------------------------*)
TYPE E_DL_HumOverrideState :
(
    eNormal         := 0,   // 正常：温控优先 / Normal, temperature control has priority
    eOverride       := 10,  // 覆盖：除湿优先生效 / Override, dehumidification has priority
    eReleasePending := 20,  // 释放待确认：湿度已回落，等确认窗 / Release pending, humidity recovered, awaiting the window
    eFault          := 99   // 故障：迟滞倒置/非有限/非法状态 / Fault, inversion, non-finite or illegal state
);
END_TYPE

FUNCTION_BLOCK FB_DL_HumidityOverride
VAR_INPUT
    fRhPct         : LREAL;                 // 实测湿度 [百分数RH] / Measured humidity [%RH]
    fRhOverridePct : LREAL := 70.0;         // 覆盖触发阈值 [百分数RH] / Override trigger threshold [%RH]
    fRhReleasePct  : LREAL := 60.0;         // 释放阈值 [百分数RH]，须 < 触发阈值 / Release threshold [%RH], must be below the trigger
    bTempCtrlActive: BOOL;                  // 温控在投 [—]（诊断参考，不参与仲裁） / Temperature control active, diagnostic reference only
    tConfirmDelay  : TIME  := T#30S;        // 触发/释放确认窗 [ms] / Trigger and release confirm window [ms]
    bReset         : BOOL;                  // 故障复位 [—] / Fault reset
END_VAR
VAR_OUTPUT
    bOverrideActive: BOOL;                  // 除湿优先生效 [—] / Dehumidification priority active
    eOverrideState : E_DL_HumOverrideState; // 仲裁相位 [—] / Arbitration phase
    eErr           : UDINT;                 // 错误码，0 = 无错 / Error code, 0 = no error
    bError         : BOOL;                  // 故障级标志，仅故障级错误置位 / Fault-class flag, set only on fault-level codes
    bValid         : BOOL;                  // 输出可用标志 / Outputs usable flag
END_VAR
VAR
    fbTrigWin      : TON;                   // 覆盖触发确认窗，段 6 无条件刷新 [ms] / Trigger confirm window
    fbReleaseWin   : TON;                   // 释放确认窗，段 6 无条件刷新 [ms] / Release confirm window
    _eState        : E_DL_HumOverrideState := E_DL_HumOverrideState.eNormal; // 当前相位 / Current phase
    _bInit         : BOOL := FALSE;         // 首扫标志，初值 FALSE 取非判定 / First-scan flag, tested negated
    _bHystBad      : BOOL;                  // 迟滞倒置/非有限锁存 / Inversion or non-finite latch
    _bSwEdge       : BOOL;                  // 切换沿单拍标志 / One-scan switch edge flag
    _bIllegal      : BOOL;                  // 非法状态标志 / Illegal state flag
END_VAR
VAR CONSTANT
    DL_HO_INF      : LREAL := 1.7976931348623157E308; // LREAL 幅值上限 / LREAL magnitude ceiling
END_VAR

(*------------------------------------------------------------------------------
 * 段 1｜每拍预置：输出先算后出，单拍标志预清零（只置必销）
 *      Outputs computed per scan, one-shot flags pre-cleared
 *-----------------------------------------------------------------------------*)
bOverrideActive := FALSE;                   // 覆盖输出每拍重算 / Override output recomputed
eErr            := 16#0000_0000;            // 错误码每拍重算 / Error code recomputed
bError          := FALSE;                   // 故障标志每拍重算 / Fault flag recomputed
bValid          := FALSE;                   // 可用标志每拍重算 / Usable flag recomputed
_bSwEdge        := FALSE;                   // 切换沿预清零 / Switch edge pre-cleared
_bIllegal       := FALSE;                   // 非法状态预清零 / Illegal flag pre-cleared

(*------------------------------------------------------------------------------
 * 段 2｜首扫初始化
 *      First-scan initialisation
 *-----------------------------------------------------------------------------*)
IF NOT _bInit THEN
    _eState   := E_DL_HumOverrideState.eNormal; // 相位正常起步 / Phase starts normal
    _bHystBad := FALSE;                     // 迟滞锁存清零 / Hysteresis latch cleared
    _bInit    := TRUE;                      // 首扫只做一次 / The first scan runs once
END_IF

(*------------------------------------------------------------------------------
 * 段 3｜组态与输入防御闸（迟滞倒置 / 湿度非有限 → 032A，保持末态）
 *      Configuration and input defense gates, last state held
 *-----------------------------------------------------------------------------*)
IF (fRhOverridePct <> fRhOverridePct) OR (ABS(fRhOverridePct) > DL_HO_INF)
   OR (fRhReleasePct <> fRhReleasePct) OR (ABS(fRhReleasePct) > DL_HO_INF) THEN
    _bHystBad := TRUE;                      // 阈值非有限归入迟滞倒置（R90） / Non-finite thresholds folded into the inversion fault
END_IF
IF (fRhPct <> fRhPct) OR (ABS(fRhPct) > DL_HO_INF) THEN
    _bHystBad := TRUE;                      // 湿度非有限：转故障态（退出覆盖由切换沿 01EE 显式声明） / Non-finite humidity, to fault, exit declared via the switch edge
END_IF
IF (NOT _bHystBad) AND (fRhReleasePct >= fRhOverridePct) THEN
    _bHystBad := TRUE;                      // 迟滞倒置锁存 / Inversion latched
END_IF
IF bReset THEN
    _bHystBad := FALSE;                     // 复位清锁存 / Reset clears the latch
END_IF

(*------------------------------------------------------------------------------
 * 段 4｜双确认窗无条件刷新（R40：CASE 之外每拍必调，各司其职不复用）
 *      Both confirm windows refreshed unconditionally per R40
 *-----------------------------------------------------------------------------*)
fbTrigWin(IN := (NOT _bHystBad) AND (_eState = E_DL_HumOverrideState.eNormal)
              AND (fRhPct >= fRhOverridePct), PT := tConfirmDelay); // 覆盖触发确认窗 / Trigger confirm window
fbReleaseWin(IN := (NOT _bHystBad) AND (_eState = E_DL_HumOverrideState.eReleasePending)
                 AND (fRhPct <= fRhReleasePct), PT := tConfirmDelay); // 释放确认窗 / Release confirm window

(*------------------------------------------------------------------------------
 * 段 5｜相位机（只做迁移；输出在段 6 按相置位）
 *      Phase machine, transitions only, outputs assigned in segment six
 *-----------------------------------------------------------------------------*)
IF _bHystBad THEN
    IF _eState <> E_DL_HumOverrideState.eFault THEN
        _bSwEdge := TRUE;                   // 进故障也按切换沿声明（画面提示） / Entering fault declared as a switch edge
    END_IF
    _eState := E_DL_HumOverrideState.eFault; // 异常转故障（保持末态由输出段承担） / Anomaly to fault
ELSE
CASE _eState OF

    E_DL_HumOverrideState.eNormal:         // 正常：触发确认窗满进覆盖
        IF fbTrigWin.Q THEN
            _bSwEdge := TRUE;               // 切换沿单发 / Switch edge one-shot
            _eState  := E_DL_HumOverrideState.eOverride; // 进覆盖 / To override
        END_IF

    E_DL_HumOverrideState.eOverride:       // 覆盖：湿度回落至释放阈进待确认
        IF fRhPct <= fRhReleasePct THEN
            _eState := E_DL_HumOverrideState.eReleasePending; // 进释放待确认 / To release pending
        END_IF

    E_DL_HumOverrideState.eReleasePending: // 释放待确认：确认窗满回正常；回弹超触发阈返覆盖
        IF fbReleaseWin.Q THEN
            _bSwEdge := TRUE;               // 切换沿单发 / Switch edge one-shot
            _eState  := E_DL_HumOverrideState.eNormal; // 回正常 / Back to normal
        ELSIF fRhPct >= fRhOverridePct THEN
            _eState := E_DL_HumOverrideState.eOverride; // 湿度回弹，返覆盖（窗自然断） / Humidity rebounded, back to override
        END_IF

    E_DL_HumOverrideState.eFault:          // 故障：复位沿且原因消失回正常
        IF bReset AND (NOT _bHystBad) THEN
            _eState := E_DL_HumOverrideState.eNormal; // 回正常 / Back to normal
        END_IF

    ELSE                                   // 非法状态兜底（R21：CASE 必带 ELSE）
        _bIllegal := TRUE;                 // 标记非法状态 / Flag the illegal state
        _eState   := E_DL_HumOverrideState.eFault; // 回故障态 / Back to fault
END_CASE
END_IF

(*------------------------------------------------------------------------------
 * 段 6｜输出置位与码位出口（职责边界：本件只仲裁，不写温度设定值）
 *      Output assignment and codes, arbitration only, no setpoint writes
 *-----------------------------------------------------------------------------*)
bOverrideActive := (_eState = E_DL_HumOverrideState.eOverride)
                OR (_eState = E_DL_HumOverrideState.eReleasePending); // 覆盖态与待确认期均视为生效 / Active in override and pending
eOverrideState := _eState;                  // 相位出口 / Phase outlet

IF _bIllegal THEN
    eErr   := 16#0005_032C;                 // 故障级：状态机兜底 / Fault: state machine fallback
    bError := TRUE;                         // 置故障标志 / Raise the fault flag
ELSIF _bHystBad THEN
    eErr   := 16#0005_032A;                 // 故障级：迟滞倒置或湿度非有限（R90 复用） / Fault: inversion or non-finite, code reused
    bError := TRUE;                         // 置故障标志 / Raise the fault flag
    bValid := FALSE;                        // 输出不可用 / Outputs unusable
ELSIF _bSwEdge THEN
    eErr := 16#0005_01EE;                   // 信息级：覆盖状态切换沿 / Info: override switch edge
    bValid := TRUE;                         // 输出可用 / Outputs usable
ELSE
    bValid := TRUE;                         // 输出可用 / Outputs usable
END_IF
END_FUNCTION_BLOCK

(* ---- FB_DL_HydronicDeltaTGuard.st ---- *)
(*
  FB_DL_HydronicDeltaTGuard  —  水系统大/小温差失衡诊断 / Hydronic delta-T imbalance diagnostic guard
  分类 Category : DL_Process
  码位 Code     : 16#06_0_94
  版本 Version  : 1.0.0
  溯源 Source   : OSCAT Building 暖通语义借鉴 · clean-room 实现，仅借分类/参数域/命名，未复制源码
  功能 Function : 1) 供/回水温差带判定：大温差（低流量征兆）/ 小温差（旁通泄漏征兆）/ 正常三档；
                  2) 旁通泄漏判据：旁通开度大且温差小持续 N 分钟（确认窗）才判泄漏；
                  3) 判据全部带迟滞防抖（回差带电平判定）。
  边界 Boundary : ① 两温度任一无效：冻结判定保持上次输出，不塞伪值；
                  ② 温差 = 0 邻域（|ΔT| < 0.5 K）判「无有效流量」而非除零算比率；
                  ③ 大/小温差判据带迟滞防抖；
                  ④ 失衡解除路径自证可达（恢复窗内即解除，泄漏需旁通关小确认）；
                  ⑤ 输出三行同向：温差档位 → 泄漏标志 → 诊断码。
  依赖 Depends  : FC_DL_Hysteresis（回差带判定，函数调用，状态由调用方持有）

  码表 Error codes（本件子码步进 16#30 · 本格 94 与既有 9X 子码段冲突，错位至 C4/D4 避让）:
    16#0002_06C4 故障级：组态非法（温差门限倒置 / 迟滞 <= 0 / 确认窗 <= 0 / 旁通门限域非法）
    16#0002_06D4 故障级：相 ID 越界（枚举兜底路径）
    16#0002_06B4 信息级：温度无效判定冻结 / 无有效流量(|ΔT|<0.5K)档（不置 bError）
*)

TYPE E_DL_HdtBand :
(
    eNormal   := 0,  // 温差正常 / Normal delta-T
    eBigDt    := 10, // 大温差（低流量征兆）/ Large delta-T, low flow sign
    eSmallDt  := 20, // 小温差（旁通泄漏征兆）/ Small delta-T, bypass leak sign
    eNoFlow   := 30, // 无有效流量（|ΔT| < 0.5 K）/ No effective flow
    eFrozen   := 40  // 温度无效冻结 / Frozen by invalid temperature
);
END_TYPE

TYPE E_DL_HdtPhase :
(
    eIdle  := 0,   // 空闲 / Idle
    eWatch := 10,  // 温差带监视 / Delta-T band watching
    eFault := 90   // 组态故障锁定 / Configuration fault locked
);
END_TYPE

FUNCTION_BLOCK FB_DL_HydronicDeltaTGuard
VAR_INPUT
    bEnable       : BOOL;                           // 总使能，FALSE 回空闲 / Master enable
    bReset        : BOOL;                           // 复位，上升沿清组态故障 / Reset, clears fault
    fSupplyC      : REAL;                           // 供水温度 [°C] / Supply water temperature [degC]
    fReturnC      : REAL;                           // 回水温度 [°C] / Return water temperature [degC]
    fBypassPct    : REAL;                           // 旁通阀开度 [%] / Bypass valve opening [%]
    fBigDtK       : REAL := 12.0;                   // 大温差门限 [K]（超过判大温差）/ Large delta-T threshold [K]
    fSmallDtK     : REAL := 4.0;                    // 小温差门限 [K]（低于判小温差）/ Small delta-T threshold [K]
    fHystK        : REAL := 1.0;                    // 迟滞回差 [K]，域 > 0 / Hysteresis band [K]
    fBypassHiPct  : REAL := 60.0;                   // 旁通开度门限 [%] / Bypass opening threshold [%]
    uLeakMin      : UINT := 10;                     // 泄漏确认窗 [min] / Leak confirm window [min]
    fTaskCycle    : REAL := 1.0;                    // 任务周期 [s]，域 > 0 / Task cycle [s]
    fEps          : REAL := 1.0E-6;                 // 浮点判零容差 [1] / Floating zero tolerance
END_VAR
VAR_OUTPUT
    eBandOut      : E_DL_HdtBand;                   // 温差档位出口 / Delta-T band output
    fDeltaTK      : REAL;                           // 当前温差 [K] / Current delta-T [K]
    bBypassLeak   : BOOL;                           // 旁通泄漏标志（确认窗后锁存）/ Bypass leak flag, latched after confirm
    bFrozen       : BOOL;                           // 判定冻结标志 / Judgment frozen flag
    bError        : BOOL;                           // 故障标志，与故障级码配对 / Fault flag
    uErrorId      : UDINT;                          // 事件码，0 = 无事件 / Event code
    eStateOut     : E_DL_HdtPhase;                  // 状态机当前态，段尾单点映射 / Phase mapped at tail
END_VAR
VAR
    _eState       : E_DL_HdtPhase := E_DL_HdtPhase.eIdle;  // 内部状态 / Internal state
    rtrReset      : R_TRIG;                         // 复位沿 / Reset edge
    bHystBig      : BOOL;                           // 大温差迟滞状态（FC_DL_Hysteresis 持有量）/ Big-delta-T hysteresis state
    bHystSmall    : BOOL;                           // 小温差迟滞状态 / Small-delta-T hysteresis state
    tonLeak       : TON;                            // 泄漏确认窗定时器 / Leak confirm window timer
    bCfgOk        : BOOL;                           // 组态合法标志 / Configuration valid
    bTempOk       : BOOL;                           // 双温度本拍有效 / Both temperatures valid
    bBypassOk     : BOOL;                           // 旁通开度本拍有效 / Bypass opening valid
    fUpInfo       : REAL;                           // 迟滞函数上阈值回读 [K] / Hysteresis upper trip readback [K]
    fLoInfo       : REAL;                           // 迟滞函数下阈值回读 [K] / Hysteresis lower trip readback [K]
    uErrH1        : UDINT;                          // 迟滞函数错误码回读 / Hysteresis error readback
    uErrH2        : UDINT;                          // 第二迟滞错误码回读 / Second hysteresis error readback
    uFault        : UDINT;                          // 锁存故障码 / Latched fault code
    uInfo         : UDINT;                          // 信息级码 / Information code
END_VAR
VAR CONSTANT
    DL_HDT_INFMAX : REAL := 1.0E30;                 // 温度有限值幅值上限 [°C] / Temperature finite bound [degC]
    DL_HDT_NOFLOW : REAL := 0.5;                    // 无有效流量邻域 [K] / No-effective-flow band [K]
END_VAR

(* === 段 0 · 实例刷新 === *)
rtrReset(CLK := bReset);                          // 每拍刷新复位沿

(* === 段 1 · 组态闸 === *)
bCfgOk := (fBigDtK > fSmallDtK + fHystK)          // 门限不倒置且迟滞带不相交
          AND (fHystK > fEps) AND (fTaskCycle > fEps)
          AND (fBypassHiPct > fEps) AND (fBypassHiPct < 100.0)   // 旁通门限域
          AND (uLeakMin >= UINT#1)                // 确认窗下限
          AND (fBigDtK = fBigDtK) AND (fSmallDtK = fSmallDtK);   // NaN 自反
IF NOT bCfgOk THEN
    uFault := 16#0002_06C4;                       // 故障级：组态非法
END_IF
IF rtrReset.Q AND bCfgOk THEN
    uFault := 16#0000;                            // 复位沿清锁存（解除路径可达）
    bBypassLeak := FALSE;                         // 泄漏标志同步复位
END_IF
uInfo := 16#0000;                                 // 信息码每拍清零
bTempOk := (fSupplyC = fSupplyC) AND (ABS(fSupplyC) < DL_HDT_INFMAX)
           AND (fReturnC = fReturnC) AND (ABS(fReturnC) < DL_HDT_INFMAX);  // 双温度 NaN 自反 + 幅值闸
bBypassOk := (fBypassPct = fBypassPct) AND (fBypassPct >= 0.0) AND (fBypassPct <= 100.0);  // 旁通域闸

(* === 段 2 · 温差折算与迟滞档位判定 === *)
fDeltaTK := 0.0;                                  // 温差缺省 0
eBandOut := E_DL_HdtBand.eFrozen;                 // 档位缺省冻结（无效时保持语义由下段覆盖）
IF bTempOk THEN
    fDeltaTK := fSupplyC - fReturnC;              // 温差 = 供 − 回 [K]
    IF ABS(fDeltaTK) < DL_HDT_NOFLOW THEN
        eBandOut := E_DL_HdtBand.eNoFlow;         // 零邻域：无有效流量档（不除零算比率）
        uInfo := 16#0002_06B4;                    // 信息级：无有效流量档
        bHystBig := FALSE;                        // 迟滞状态同步复位
        bHystSmall := FALSE;
    ELSE
        FC_DL_Hysteresis(fIn := fDeltaTK,         // 大温差迟滞判定（状态由本件持有）
                         fThreshold := fBigDtK,   // 设定点 = 大温差门限
                         fHysteresis := fHystK,   // 回差带
                         bState := bHystBig,      // 持有状态回传（IN_OUT）
                         fUpperTrip => fUpInfo, fLowerTrip => fLoInfo,
                         uErrorId => uErrH1);     // 输出取值用 => 显式接收
        FC_DL_Hysteresis(fIn := fDeltaTK,         // 小温差迟滞判定
                         fThreshold := fSmallDtK,
                         fHysteresis := fHystK,
                         bState := bHystSmall,
                         fUpperTrip => fUpInfo, fLowerTrip => fLoInfo,
                         uErrorId => uErrH2);
        IF bHystBig THEN
            eBandOut := E_DL_HdtBand.eBigDt;      // 大温差档（回差带内保持，防抖）
        ELSIF bHystSmall THEN
            eBandOut := E_DL_HdtBand.eSmallDt;    // 小温差档
        ELSE
            eBandOut := E_DL_HdtBand.eNormal;     // 正常档
        END_IF
    END_IF
ELSE
    (* 温度无效：保持上次档位输出（不塞伪值，冻结标志由段尾映射） *)
    uInfo := 16#0002_06B4;                        // 信息级：温度无效判定冻结
END_IF

(* === 段 3 · 旁通泄漏确认窗（泄漏需持续 N 分钟才判）=== *)
tonLeak(IN := bTempOk AND bBypassOk AND (eBandOut = E_DL_HdtBand.eSmallDt)
             AND (fBypassPct >= fBypassHiPct),    // 小温差 + 旁通大开度同时成立才计时
        PT := REAL_TO_TIME(UINT_TO_REAL(uLeakMin) * 60.0 * 1000.0));   // 确认窗换算 [ms]（UINT 扩宽 REAL 防溢出）
IF tonLeak.Q THEN
    bBypassLeak := TRUE;                          // 确认窗满：泄漏锁存
END_IF
IF bTempOk AND bBypassOk AND ((eBandOut = E_DL_HdtBand.eNormal)
    OR (eBandOut = E_DL_HdtBand.eBigDt) OR (fBypassPct < fBypassHiPct - fEps)) THEN
    bBypassLeak := FALSE;                         // 恢复正常档或旁通关小：解除（路径可达）
END_IF

(* === 段 4 · 主状态机（ENUM + CASE，含 ELSE 兜底）=== *)
CASE _eState OF
E_DL_HdtPhase.eIdle :
    IF uFault <> 16#0000 THEN
        _eState := E_DL_HdtPhase.eFault;          // 故障优先
    ELSIF bEnable AND bCfgOk THEN
        _eState := E_DL_HdtPhase.eWatch;          // 进监视相
    END_IF

E_DL_HdtPhase.eWatch :
    IF (uFault <> 16#0000) OR (NOT bEnable) THEN
        _eState := E_DL_HdtPhase.eFault;          // 故障/失能转出
    END_IF

E_DL_HdtPhase.eFault :
    IF uFault = 16#0000 THEN
        _eState := E_DL_HdtPhase.eIdle;           // 解锁回空闲
    END_IF

ELSE
    _eState := E_DL_HdtPhase.eFault;              // 非法状态拦截
    uFault := 16#0002_06D4;                       // 故障级：相 ID 越界
END_CASE
bFrozen := (NOT bTempOk) OR (_eState = E_DL_HdtPhase.eFault);   // 冻结标志段尾单点映射

(* === 段 5 · 输出映射 === *)
bError := (uFault <> 16#0000);                    // 故障标志仅由故障级码置位（R45 配对）
IF bError THEN
    uErrorId := uFault;                           // 故障级优先上报
ELSE
    uErrorId := uInfo;                            // 否则上报信息级码
END_IF
eStateOut := _eState;                             // 输出枚举段尾单点映射（N2 规则）
END_FUNCTION_BLOCK

(* ---- FB_DL_HydronicMeterAudit.st ---- *)
(*
  FB_DL_HydronicMeterAudit  —  冷冻水/冷却水能量审计（流量累计 × 侧焓差） / Hydronic energy audit: flow accumulation times loop enthalpy difference
  分类 Category : DL_Process
  版本 Version  : 1.0.1
  来源 Source   : t1-2-oscat-building — 楼宇能量审计族零检索深化
  溯源 Origin   : clean-room 实现，Q = 流量×密度×比热×温差 换算链为公开热工公式，未复制任何源码行
  功能 Function : 1) 逐周期功率换算：fPowerKw = fFlowLpm × fRhoKgL × fCpKj ×
                  (fTinC - fToutC) / 60.0（L/min×kg/L×kJ/(kg·K)×K = kJ/min，
                  除以 60 得 kW，除数 60.0 为常量无除零）；
                  2) 能量累计：fEnergyKwh += fPowerKw × tCycle/T#1H（TIME 比
                  经 DINT 除法，除数 T#1H 为非零常量）；累计仅使能相且温差判据
                  有效（|ΔT| >= fDtMinK）承载；
                  3) 温差判据无效（|ΔT| < fDtMinK）→ ePause 相暂停累计（ePause
                  双出口：判据恢复 / 撤使能，R98）；累计饱和（fEnergyKwh 越上限
                  1.0E12，可表性反算：远低于 LREAL 上限 1.8E308）→ 0387 锁存；
                  4) 故障级：0385 组态非法 / 0386 输入非有限锁存 / 0387 饱和锁存；
                  5) 信息级三码：审计激活沿 / 温差判据恢复沿 / 累计复位完成沿；
                  6) 解除式全当拍量（R240 落地），逐 BOOL 标注见段 4。
  边界 Boundary : ① 组态闸：tCycle <= 0、fCpKj <= 0、fRhoKgL <= 0、fDtMinK < 0
                  → 0385 锁存，ELSE 兜底归并 0385（码表声明），累计停发；
                  ② 非有限判据用自反比较与差值自减双判（禁近似阈值，R79）；
                  ③ ΔT 上下双向均参与功率（冷/热侧同式），不按方向拆分归因
                  （本件为能量计量非保护判据，R146 方向拆分不适用）；
                  ④ 无 GVL 依赖：纯引脚输入输出，无外部变量引用，无物理 IO 地址。
  依赖 Depends  : Standard.library（TON / R_TRIG）
  码表 Error codes（Process 段 0005，窗口 0385~0387 / 04AD~04AF）:
    16#0005_0385 故障级：组态非法（周期/比热/密度/温差阈域非法）或相位落 ELSE 兜底（归并声明），锁存至 bReset
    16#0005_0386 故障级：流量或温度输入非有限锁存（累计暂停，安全侧），锁存至 bReset
    16#0005_0387 故障级：能量累计饱和锁存（越 1.0E12 kWh 上限，停止累计），锁存至 bReset
    16#0005_04AD 信息级：审计激活沿（进 eRun）
    16#0005_04AE 信息级：温差判据恢复沿（ePause 判据恢复出口）
    16#0005_04AF 信息级：能量累计复位完成沿
  修订历史 Revision :
    2026-11-19  v1.0.0  R42 首版（批次 2 · 序号 3）
    2026-11-19  v1.0.1  R42 终审返修：① 补声明内部相位变量 _eState（首版漏声明，
                        段 4/CASE 引用未声明变量属编译阻断缺陷，机检盲区）；
                        ② 新增段 4A 故障锁存相位迁移闸——0385/0386/0387 锁存后
                        _eState 强制迁 eFault，冻结 eRun 相内累计递增（否则饱和
                        锁存后 fEnergyKwh 持续越限增长、0385 期间累计不冻结）；
                        对外引脚契约不变。
*)

TYPE E_DL_HmaState :
(
    eIdle   := 0,    // 未使能：不累计 / Idle, not accumulating
    eRun    := 10,   // 审计中：逐周期累计 / Run, per-cycle accumulating
    ePause  := 20,   // 暂停：温差判据无效 / Pause, delta-T verdict invalid
    eFault  := 90    // 故障：非有限或饱和锁定 / Fault, latched
);
END_TYPE

FUNCTION_BLOCK FB_DL_HydronicMeterAudit
VAR_INPUT
    fFlowLpm     : REAL := 0.0;       // 侧流量 [L/min]，调用方注入 / Loop flow rate
    fTinC        : REAL := 12.0;      // 供水温度 [°C] / Supply water temperature
    fToutC       : REAL := 7.0;       // 回水温度 [°C] / Return water temperature
    fCpKj        : REAL := 4.186;     // 水比热 [kJ/(kg·K)]，域 > 0 / Specific heat capacity
    fRhoKgL      : REAL := 1.0;       // 水密度 [kg/L]，域 > 0 / Water density
    fDtMinK      : REAL := 0.5;       // 温差判据下限 [K]，域 >= 0 / Minimum delta-T verdict threshold
    fEnergyCap   : REAL := 1.0E12;    // 能量累计上限 [kWh]，可表性反算见头注释 / Energy accumulation cap
    tCycle       : TIME := T#1S;      // 审计累加周期 [ms]，域 > 0 / Audit accumulation cycle
    bAuditEn     : BOOL := FALSE;     // 审计使能（电平）[-] / Audit enable, level
    bEnergyRst   : BOOL := FALSE;     // 能量复位指令，上升沿清累计 [-] / Energy reset command edge
    bReset       : BOOL := FALSE;     // 复位，上升沿清故障锁存 / Reset edge clears fault latch
END_VAR
VAR_OUTPUT
    eState       : E_DL_HmaState;     // 状态出口，段尾单点映射 / State outlet
    fPowerKw     : REAL;              // 逐周期功率 [kW] / Per-cycle power
    fEnergyKwh   : REAL;              // 能量累计 [kWh] / Accumulated energy
    bDtInvalid   : BOOL;              // 温差判据无效镜像 [-] / Delta-T invalid mirror
    bError       : BOOL;              // 故障锁存标志 / Fault latch flag
    nErrId       : UDINT;             // 事件码，0 = 无事件 / Event code
END_VAR
VAR
    _eState      : E_DL_HmaState := E_DL_HmaState.eIdle;  // 内部相位（CASE 唯一写入目标；R42 终审补声明）/ Internal phase
    rtEnergyRst  : R_TRIG;            // 能量复位沿实例，无条件刷新 / Energy reset edge instance
    rtReset      : R_TRIG;            // 复位沿实例，无条件刷新 / Reset edge instance
    _fDt         : REAL;              // 侧温差 [K]（当拍量）/ Loop delta temperature
    _bDtOk       : BOOL;              // 温差判据有效当拍量 [-] / Delta-T verdict valid flag
    _bNonFin     : BOOL;              // 输入非有限当拍量 [-] / Non-finite input flag
    _bFault      : BOOL;              // 故障锁存位（锁存量）/ Latched fault bit
    _uFault      : UDINT;             // 故障码锁存（锁存量）/ Latched fault code
    _uInfo       : UDINT;             // 信息码，每拍重算 / Transient info code
END_VAR

(* —— 段 0：沿实例无条件周期刷新（禁置于 IF/CASE 内） —— *)
_fDt := fTinC - fToutC;                              // 侧温差（当拍量）
_bDtOk := ABS(_fDt) >= fDtMinK;                      // 温差判据有效（当拍量，容差式阈值）
_bNonFin := (fFlowLpm <> fFlowLpm) OR (fTinC <> fTinC) OR (fToutC <> fToutC)
         OR ((fFlowLpm - fFlowLpm) <> (fFlowLpm - fFlowLpm))
         OR ((fTinC - fTinC) <> (fTinC - fTinC))
         OR ((fToutC - fToutC) <> (fToutC - fToutC));        // 非有限防御（NaN 自反 + 差值自减）
rtEnergyRst(CLK := bEnergyRst);                      // 能量复位沿（每拍必调）
rtReset(CLK := bReset);                              // 复位沿（每拍必调）

(* —— 段 1：单拍量预清零（锁存量 _bFault/_uFault 不入清单，禁同拍抹除） —— *)
_uInfo := 16#0000_0000;             // 信息码每拍重算
fPowerKw := 0.0;                    // 功率出口缺省 0
bDtInvalid := FALSE;                // 判据无效镜像缺省 FALSE
nErrId := 16#0000_0000;             // 事件码缺省无事件

(* —— 段 2：复位沿 + 组态域闸（当拍量判据） —— *)
IF rtReset.Q THEN                   // rtReset.Q = 当拍量
    _bFault := FALSE;               // 清故障锁存位
    _uFault := 16#0000_0000;        // 清故障锁存码
END_IF
IF (TIME_TO_DINT(tCycle) <= 0) OR (fCpKj <= 0.0) OR (fRhoKgL <= 0.0) OR (fDtMinK < 0.0) THEN
    _uFault := 16#0005_0385;        // 故障级：组态非法
    _bFault := TRUE;                // 故障标志与码位配对（R45）
END_IF
IF rtEnergyRst.Q THEN               // 能量复位沿（当拍量）
    fEnergyKwh := 0.0;              // 累计清零
    _uInfo := 16#0005_04AF;         // 信息级：累计复位完成沿
END_IF

(* —— 段 3：非有限与饱和锁存（判据当拍量；安全侧赋值右值仅常量，FB32-4） —— *)
IF _bNonFin THEN
    fPowerKw := 0.0;                // 安全侧功率清零（常量右值）
    _uFault := 16#0005_0386;        // 故障级：输入非有限锁存
    _bFault := TRUE;
END_IF
IF (NOT _bFault) AND (fEnergyKwh >= fEnergyCap) THEN
    _uFault := 16#0005_0387;        // 故障级：累计饱和锁存
    _bFault := TRUE;
END_IF

(* —— 段 4：故障解除式（R240 落地，逐 BOOL 标注）：
     rtReset.Q = 当拍量；NOT _bNonFin = 当拍量；NOT bAuditEn = 当拍量；
     fEnergyKwh < fEnergyCap 为保持槽值（非当拍量），饱和解除路径为能量复位沿 + 复位沿组合：
     rtEnergyRst.Q 先清 fEnergyKwh，下一拍保持槽值已降，复位沿当拍量配合解除。 —— *)
IF rtReset.Q AND (NOT _bNonFin) AND (NOT bAuditEn) THEN
    _bFault := FALSE;               // 清故障锁存位（锁存量，仅此当拍量解除沿可清）
    _uFault := 16#0000_0000;        // 清故障锁存码（锁存量，仅本当拍量解除沿可清）
    IF _eState = E_DL_HmaState.eFault THEN
        _eState := E_DL_HmaState.eIdle;     // 故障相迁出：回未使能
    END_IF
END_IF

(* —— 段 4A：故障锁存相位迁移闸（R42 终审返修，v1.0.1）：
     0385 组态 / 0386 非有限 / 0387 饱和锁存置位而相位未迁出时强制入故障相，
     冻结 eRun 相内累计递增（否则饱和锁存后 fEnergyKwh 每周期持续越限增长，
     0385 组态非法期间累计亦不冻结）；置于段 4 之后，解除沿当拍清锁不触发
     迁移，无同拍抢迁。 —— *)
IF _bFault AND (_eState <> E_DL_HmaState.eFault) THEN
    _eState := E_DL_HmaState.eFault;        // 锁存即入故障相（累计冻结，仅解除沿可离相）
END_IF

(* —— 段 5：相位机（CASE 全覆盖 + ELSE 兜底；累计仅在段内承载） —— *)
CASE _eState OF

E_DL_HmaState.eIdle:
    IF bAuditEn AND (NOT _bFault) THEN
        _uInfo := 16#0005_04AD;         // 信息级：审计激活沿
        _eState := E_DL_HmaState.eRun;  // 进审计相
    END_IF

E_DL_HmaState.eRun:
    IF (NOT _bNonFin) AND _bDtOk THEN   // 判据有效：逐周期累计（除数 60.0/T#1H 均非零常量）
        fPowerKw := (LREAL_TO_REAL(LREAL(fFlowLpm) * LREAL(fRhoKgL) * LREAL(fCpKj)
                    * LREAL(_fDt) / 60.0));         // 功率换算（LREAL 精度承载）
        fEnergyKwh := fEnergyKwh + fPowerKw * LREAL_TO_REAL(TIME_TO_LREAL(tCycle) / TIME_TO_LREAL(T#1H));
                                        // 能量累计（周期占比加权）
    ELSE
        _eState := E_DL_HmaState.ePause;    // 判据无效：进暂停相
    END_IF
    IF NOT bAuditEn THEN
        _eState := E_DL_HmaState.eIdle;     // 撤使能：回未使能相
    END_IF

E_DL_HmaState.ePause:
    bDtInvalid := TRUE;                 // 判据无效镜像（相电平）
    IF _bDtOk AND (NOT _bNonFin) THEN   // 出口 1：判据恢复（事件量）
        _uInfo := 16#0005_04AE;         // 信息级：温差判据恢复沿
        _eState := E_DL_HmaState.eRun;  // 回审计相
    ELSIF NOT bAuditEn THEN             // 出口 2：撤使能（前置条件消失，R98 双出口）
        _eState := E_DL_HmaState.eIdle; // 回未使能相
    END_IF

E_DL_HmaState.eFault:
    ;                                   // 故障相：累计冻结，等解除沿（段 4 承载迁出）

ELSE
    _uFault := 16#0005_0385;            // 故障级：非法相位兜底（归并组态码，码表声明）
    _bFault := TRUE;
    _eState := E_DL_HmaState.eFault;    // 强制回故障相

END_CASE

(* —— 段 6：出口单点映射（名实同源；锁存码回放，禁同拍抹除） —— *)
IF _bFault THEN
    nErrId := _uFault;              // 故障锁存码回放
    fPowerKw := 0.0;                // 故障相功率出口强制 0（安全侧）
    bDtInvalid := FALSE;            // 故障相判据镜像强制 FALSE
ELSE
    nErrId := _uInfo;               // 信息码
END_IF
bError := _bFault;                  // 故障标志与锁存位同源
eState := _eState;                  // 状态出口单点映射

END_FUNCTION_BLOCK

(* ---- FB_DL_HydrostaticLevelComp.st ---- *)
(*==============================================================================
 * 组件名称 (Component)  : FB_DL_HydrostaticLevelComp
 * 所属子库 (Sublibrary) : DL_Process
 * 前缀     (Prefix)     : FB_DL_
 * 当前版本 (Version)    : 1.0.0
 * 兼容性   (Platform)   : CODESYS 3.5 / TwinCAT 3 / 汇川 InoProShop / Schneider
 *                         Machine Expert；纯 IEC 61131-3（第 3 版），
 *                         仅依赖标准库 R_TRIG / ABS / MAX / MIN 与库内
 *                         FC_DL_MultiPointLinear（分段线性插值复用），
 *                         零厂商方言
 * 作者     (Author)     : 道莅代码库 · PLC编程专家（R31）
 * 开源溯源 (Origin)     : 静压式液位计介质密度温补公开工艺语义（行业池），
 *                         道莅 clean-room 防御性实现，未复制任何外部源码行
 * 功能描述 (Function)   : 静压液位介质密度温补件。介质密度由温度-密度标定表
 *                         经库内 FC_DL_MultiPointLinear 分段线性插值得到；
 *                         液位 = (压强 − 干扰管偏移) / (密度 × g)，重力加速度
 *                         g = 9.80665 米每二次方秒常量写死本头注释；表外
 *                         温度最近端点钳位记信息码。密度单位 千克每立方米、
 *                         液位单位 米 必标。
 * 依赖表   (Depends)    : FC_DL_MultiPointLinear（折线插值，IN-OUT 数组注入）。
 * 码位     (Codes)      : 16#0005_00C1 信息级：温度表外钳位照算（不置 bError）
 *                         16#0005_00C2 故障级：密度退化（插值结果不大于
 *                                      1E-6 拒算早退）与输入非有限
 *                         16#0005_00C3 故障级：标定表非单调（锁存）
 *                         16#0005_00C4 故障级：标定表空/点数不足（锁存）
 *                         16#0005_00C5 保留未启用（码表与实现对齐）
 * 边界防错 (Boundary)   : 1 密度不大于 1.0E-6 拒算早退防除零；
 *                         2 非有限全拦（x<>x 自反判加幅值界）；
 *                         3 标定表须严格递增否则组态码锁存；
 *                         4 表点数 0/1 组态非法（故障级锁存）；
 *                         5 故障锁存可达解除路径：bRst 复位沿；
 *                         6 R_TRIG 实例每拍无条件刷新。
 * 修订历史 (Revision)   : 2026-11-18 v1.0.0 首版入库（R31 · 阶段三 · 序 19）
 *==============================================================================*)

(*------------------------------------------------------------------------------
 * 结构体: ST_DL_Pt2（归属本功能块，同文件发布，全库唯一属主）
 *----------------------------------------------------------------------------*)
TYPE ST_DL_Pt2 :
STRUCT
    fX : REAL := 0.0;   // 折点自变量：温度 [摄氏度] / Breakpoint X: temperature [degC]
    fY : REAL := 0.0;   // 折点因变量：密度 [千克每立方米] / Breakpoint Y: density [kg per m3]
END_STRUCT
END_TYPE

(*==============================================================================
 * 功能块: FB_DL_HydrostaticLevelComp
 * 调用约定: 每个扫描周期无条件调用一次；标定表经引脚数组注入（上限 16 点）。
 *==============================================================================*)
FUNCTION_BLOCK FB_DL_HydrostaticLevelComp
VAR_INPUT
    fPMeas  : REAL := 0.0;            // 静压压强实测 [千帕] / Measured hydrostatic pressure [kPa]
    fTCurve : ARRAY[1..16] OF ST_DL_Pt2; // 温度-密度标定表 [摄氏度-千克每立方米] / Temperature-density calibration table
    uPtCnt  : UINT := 16;             // 有效标定点数 [个]，合法域 2..16 / Valid point count, valid 2..16
    fTNow   : REAL := 20.0;           // 介质温度实测 [摄氏度] / Medium temperature [degC]
    fDpOffset: REAL := 0.0;           // 干扰管偏移 [千帕] / Dry-leg offset [kPa]
    bEn     : BOOL := FALSE;          // 使能 / Enable flag
    bRst    : BOOL := FALSE;          // 组态故障复位沿（可增引脚）/ Config fault reset edge, added pin
END_VAR
VAR_OUTPUT
    fLevel  : REAL;                   // 补偿后液位 [米] / Compensated level [m]
    fDensity: REAL;                   // 介质密度 [千克每立方米] / Medium density [kg per m3]
    bValid  : BOOL;                   // 输出可用标志 / Output validity flag
    bError  : BOOL;                   // 故障标志 / Error flag
    uErrorId: UDINT;                  // 错误码，0 = 无错 / Error code, 0 = none
END_VAR
VAR
    rTrigRst: R_TRIG;                 // 复位沿检测，每拍无条件刷新 / Reset edge detector, refreshed every scan
    afX     : ARRAY[0..15] OF LREAL;  // 插值件自变量表 [摄氏度] / Interpolation X table [degC]
    afY     : ARRAY[0..15] OF LREAL;  // 插值件因变量表 [千克每立方米] / Interpolation Y table [kg per m3]
    bClamped: BOOL;                   // 插值钳位标志 / Interpolation clamp flag
    bExtra  : BOOL;                   // 插值外推标志 / Interpolation extrapolation flag
    nSeg    : INT;                    // 插值命中段号 / Interpolation segment index
    uErrMPL : UDINT;                  // 插值件错误码 / Interpolation error code
    nCntEff : INT;                    // 钳位后点数 [个] / Effective point count
    bMonoOk : BOOL;                   // 表单调标志 / Table monotonic flag
    bCntOk  : BOOL;                   // 点数合法标志 / Point count legality flag
    bInOk   : BOOL;                   // 输入有效性 / Input validity flag
    fRhoL   : LREAL;                  // 插值密度（LREAL 域）[千克每立方米] / Interpolated density [kg per m3]
    fNum    : REAL;                   // 液位分子暂存 [千帕] / Level numerator staging [kPa]
    fDen    : REAL;                   // 液位分母暂存 [千帕每米] / Level denominator staging [kPa per m]
    bCfgLatch: BOOL;                  // 组态故障锁存标志 / Config fault latch flag
    uCfgCode: UDINT;                  // 组态锁存码 / Config latched code
    i       : INT;                    // 表装载循环索引 / Table load loop index
    bClampInfo: BOOL;                 // 温度钳位信息 / Temperature clamp info flag
END_VAR
VAR CONSTANT
    DL_HLC_PT_MAX : INT   := 16;      // 标定表点数上限 [个] / Calibration point upper bound
    DL_HLC_FIN    : REAL  := 1.0E30;  // REAL 有限幅值判界 / REAL finiteness magnitude bound
    DL_HLC_G      : REAL  := 9.80665; // 重力加速度常量 [米每二次方秒]，写死头注释 / Gravity constant [m per s2], fixed in header
    DL_HLC_EPS    : REAL  := 1.0E-6;  // 密度拒算下限 [千克每立方米] / Density rejection floor [kg per m3]
    DL_HLC_KPA    : REAL  := 1000.0;  // 千帕到帕换算系数 / kPa to Pa factor
END_VAR

// ---- 段 1｜边沿实例无条件刷新（红线：禁入条件分支）----------------------------
rTrigRst(CLK := bRst);                                // 复位沿检测 / Reset edge detection

// ---- 段 2｜组态校验（点数与单调性），故障锁存带可达复位通道 ----------------------
IF rTrigRst.Q THEN
    bCfgLatch := FALSE;                               // 复位清组态锁存 / Reset clears config latch
    uCfgCode := 16#0000_0000;                         // 清锁存码 / Clear latched code
END_IF
nCntEff := MIN(UINT_TO_INT(uPtCnt), DL_HLC_PT_MAX);   // 点数钳上限 / Clamp point count
bCntOk := (nCntEff >= 2);                             // 点数 0/1 组态非法 / Point count 0 or 1 illegal
bMonoOk := TRUE;                                      // 单调标志预置 / Preset monotonic
IF bCntOk THEN
    FOR i := 1 TO (nCntEff - 1) DO
        IF (fTCurve[i].fX <> fTCurve[i].fX) OR (fTCurve[i + 1].fX <> fTCurve[i + 1].fX)
           OR (fTCurve[i + 1].fX <= fTCurve[i].fX) THEN
            bMonoOk := FALSE;                         // 非严格递增判非单调 / Non-strict increase is non-monotonic
        END_IF
    END_FOR
END_IF
IF bCntOk AND bMonoOk THEN
    bCfgLatch := FALSE;                               // 组态自愈（表改好自动解除）/ Config self-heals
    uCfgCode := 16#0000_0000;                         // 清锁存码 / Clear latched code
ELSE
    IF NOT bCntOk THEN
        uCfgCode := 16#0005_00C4;                     // 码位：表空/点数不足 / Code: table empty
    ELSE
        uCfgCode := 16#0005_00C3;                     // 码位：表非单调 / Code: table non-monotonic
    END_IF
    bCfgLatch := TRUE;                                // 组态故障锁存 / Config fault latched
END_IF

// ---- 段 3｜组态合法时装载插值表并调库内折线件（IN-OUT 数组注入）------------------
bValid := FALSE;                                      // 可用标志先清 / Clear validity
IF bCfgLatch = FALSE THEN
    FOR i := 1 TO nCntEff DO
        afX[i - 1] := REAL_TO_LREAL(fTCurve[i].fX);   // 自变量装载 / Load X table
        afY[i - 1] := REAL_TO_LREAL(fTCurve[i].fY);   // 因变量装载 / Load Y table
    END_FOR
    fRhoL := FC_DL_MultiPointLinear(afX, afY,
             fIn := REAL_TO_LREAL(fTNow), nCount := nCntEff, bClamp := TRUE,
             nSegment => nSeg, bExtrapolated => bExtra, bClamped => bClamped,
             uErrorId => uErrMPL);                    // 库内折线插值取密度 / Library interpolation for density
    fDensity := LREAL_TO_REAL(fRhoL);                 // 密度落地 [千克每立方米] / Density to REAL
    bClampInfo := bClamped;                           // 表外温度钳位信息 / Temperature clamp info
END_IF

// ---- 段 4｜液位换算（非有限全拦，密度下限拒算防除零）----------------------------
bInOk := (fPMeas = fPMeas) AND (fTNow = fTNow) AND (fDpOffset = fDpOffset)
     AND (ABS(fPMeas) < DL_HLC_FIN) AND (ABS(fTNow) < DL_HLC_FIN)
     AND (ABS(fDpOffset) < DL_HLC_FIN);               // 三输入有限 / Three inputs finite
IF bCfgLatch = FALSE THEN
    IF NOT bInOk THEN
        bValid := FALSE;                              // 非有限拒输出 / Non-finite rejects output
        uErrorId := 16#0005_00C2;                     // 故障级：输入非有限 / Fault: non-finite input
    ELSIF fDensity <= DL_HLC_EPS THEN
        bValid := FALSE;                              // 密度退化拒算早退 / Degenerate density rejects
        uErrorId := 16#0005_00C2;                     // 故障级：密度退化 / Fault: density degenerate
    ELSE
        fNum := (fPMeas - fDpOffset) * DL_HLC_KPA;    // 分子换帕 [帕] / Numerator to Pa
        fDen := fDensity * DL_HLC_G / DL_HLC_KPA;     // 分母千帕每米 [千帕每米] / Denominator kPa per m
        fLevel := fNum / fDen;                        // 液位 [米]，分母已验正 / Level [m], denominator verified
        bValid := TRUE;                               // 输出可用 / Output valid
        IF bClampInfo THEN
            uErrorId := 16#0005_00C1;                 // 信息级：温度表外钳位 / Info: temperature clamped
        ELSE
            uErrorId := 16#0000_0000;                 // 无码 / No code
        END_IF
    END_IF
END_IF

// ---- 段 5｜组态锁存回放（故障级配对置位）----------------------------------------
IF bCfgLatch THEN
    bValid  := FALSE;                                 // 组态故障拒输出 / Config fault rejects output
    bError  := TRUE;                                  // 故障标志配对（R45）/ Fault flag paired
    uErrorId := uCfgCode;                             // 锁存码回放 / Latched code replayed
ELSE
    bError := (uErrorId = 16#0005_00C2);              // 仅数值故障级置故障标志 / Only numeric fault sets flag
END_IF
END_FUNCTION_BLOCK

(* ---- FB_DL_InjectionMoldClampSeq.st ---- *)
(*
  道莅工业代码库 | DL_Process | FB_DL_InjectionMoldClampSeq
  版本: 1.0.0 | 日期: 2026-11-23 | 轮次: R75
  开源溯源: self-cleanroom（无外部来源；行业池·塑机工艺通用语义，零代码行复制）
  功能: 注塑机五段工艺序列——低压护模→高压锁模→射胶→保压→冷却→开模；
        锁模力段间闸（高压锁模后须实测力达下限才放行射胶）与护模/锁模/
        射胶/开模超时出口；中止命令走开模安全撤离（不置故障不计数）。
  兼容性: CODESYS 3.5 / TwinCAT 3 / 汇川 InoProShop；仅依赖标准 TON / R_TRIG，零厂商私有库
  接口: 输入启动/限位/实测力/实测射压/熔胶到位/各段定时/中止/复位；输出各段
        驱动输出、循环完成单拍、循环计数、eState/eCause/bError/nErrId。
  码表: 16#0005_03B7 故障级：合模序列故障总码（锁存至复位沿，归由 eCause）
        16#0005_04DA 信息级：循环完成台账（eDone 相单拍，uCycleCnt 定稿）
        16#0005_04DB 信息级：中止撤离完成（eOpen 相开到位，不计数）
        码段说明：0005 段故障子带 03xx / 信息子带 04xx，槽位经全库实扫空闲。
  边界: ① 锁模力闸：bMoldClosedLim 已到位而 fClampForceAct 低于下限 →
        等待 tForceGateWait，超时判闸失败（eCause eForceGateTimeout）；
        ② 实测力/射压 NaN 时比较恒 FALSE → 挂等待窗，超时走对应故障出口
        （NaN 不穿透段间闸，结构性防御）；
        ③ ①完成脉冲经 rtDone R_TRIG 单拍化（内部状态置位 → 统一出口映射单拍）；
        ④ 八个 TON + 三个 R_TRIG 段 0 无条件周期刷新；
        ⑤ 故障解除唯一路径 = bReset 上升沿 ∧ 组态合法；⑥ 零全局耦合。
  邻件比对: PileClampCtrl（打桩夹桩，行业域不同），无注塑合模属主（R75 §3 留痕）。
  修订历史: 2026-11-23 v1.0.0 R75 首版（复杂件批 B1 · C02）
*)

TYPE E_DL_IcsPhase :
(
    eIdle      := 0,   // 待机 | Idle
    eClampLp   := 10,  // 低压护模 | Low-pressure mold protect
    eClampHp   := 20,  // 高压锁模 | High-pressure clamp
    eInject    := 30,  // 射胶 | Injection
    eHold      := 40,  // 保压 | Packing hold
    eCool      := 50,  // 冷却 | Cooling
    eOpen      := 60,  // 开模 | Mold open
    eDone      := 70,  // 循环完成单拍相 | Cycle done one-shot phase
    eFault     := 90   // 故障锁存相 | Fault latch phase
);
END_TYPE

TYPE E_DL_IcsCause :
(
    eNone            := 0,  // 无故障 | No cause
    eCfgIllegal      := 1,  // 组态非法 | Illegal configuration
    eClampLpTimeout  := 2,  // 低压护模超时 | Low-pressure protect timeout
    eClampHpTimeout  := 3,  // 高压锁模超时 | High-pressure clamp timeout
    eForceGateTimeout:= 4,  // 锁模力段间闸等待超时 | Clamp force gate wait timeout
    eInjectTimeout   := 5,  // 射胶（含熔胶等待）超时 | Injection incl melt wait timeout
    eOpenTimeout     := 6   // 开模超时 | Mold open timeout
);
END_TYPE

FUNCTION_BLOCK FB_DL_InjectionMoldClampSeq
VAR_INPUT
    bStartCmd       : BOOL := FALSE;   // 循环启动命令（电平）[-] | Cycle start command level
    bMoldClosedLim  : BOOL := FALSE;   // 模具合到位限位 [-] | Mold closed limit switch
    bMoldOpenLim    : BOOL := FALSE;   // 模具开到位限位 [-] | Mold open limit switch
    fClampForceAct  : REAL := 0.0;     // 实测锁模力 [kN] | Actual clamp force
    fClampForceMin  : REAL := 500.0;   // 锁模力段间闸下限，域 > 0 [kN] | Clamp force gate threshold
    bMeltReady      : BOOL := FALSE;   // 熔胶计量到位（射胶前置）[-] | Melt metering ready precondition
    fInjPressAct    : REAL := 0.0;     // 实测射胶压力 [bar] | Actual injection pressure
    fInjPressSp     : REAL := 800.0;   // 射胶压力切换点设定，域 > 0 [bar] | Injection switchover pressure setpoint
    tClampLpTimeout : TIME := T#10S;   // 低压护模允许时长，域 > T#0S | LP protect allow time
    tClampHpTimeout : TIME := T#5S;    // 高压锁模允许时长，域 > T#0S | HP clamp allow time
    tForceGateWait  : TIME := T#5S;    // 锁模力闸等待超时，域 > T#0S | Force gate wait timeout
    tInjectTimeout  : TIME := T#15S;   // 射胶允许时长，域 > T#0S | Injection allow time
    tHoldTime       : TIME := T#8S;    // 保压时长，域 > T#0S | Hold duration
    tCoolTime       : TIME := T#30S;   // 冷却时长，域 > T#0S | Cooling duration
    tOpenTimeout    : TIME := T#15S;   // 开模允许时长，域 > T#0S | Open allow time
    bCycleAbort     : BOOL := FALSE;   // 循环中止命令（电平）[-] | Cycle abort command level
    bReset          : BOOL := FALSE;   // 复位命令，上升沿清故障 [-] | Reset command, rising edge
END_VAR
VAR_OUTPUT
    bClampFwd  : BOOL;                 // 合模输出（低压+高压段）[-] | Clamp forward output
    bClampHigh : BOOL;                 // 高压锁模输出 [-] | High-pressure clamp output
    bInjectOut : BOOL;                 // 射胶输出 [-] | Injection output
    bHoldOut   : BOOL;                 // 保压输出 [-] | Hold output
    bCoolOut   : BOOL;                 // 冷却输出 [-] | Cooling output
    bOpenOut   : BOOL;                 // 开模输出 [-] | Open output
    bCycleDone : BOOL;                 // 循环完成单拍脉冲 [-] | Cycle done one-shot pulse
    uCycleCnt  : UDINT;                // 完成循环计数 [次] | Completed cycle count
    eState     : E_DL_IcsPhase;        // 相位出口 | Phase outlet
    eCause     : E_DL_IcsCause;        // 故障成因出口 | Fault cause outlet
    bError     : BOOL;                 // 故障锁存标志 [-] | Fault latch flag
    nErrId     : UDINT;                // 事件码，0 = 无事件 | Event code, 0 = none
END_VAR
VAR
    _eState    : E_DL_IcsPhase := E_DL_IcsPhase.eIdle;    // 内部相位（CASE 唯一写入目标） | Internal phase
    _eCause    : E_DL_IcsCause := E_DL_IcsCause.eNone;    // 成因锁存 | Latched cause
    _bFault    : BOOL;                 // 故障锁存位 | Fault latch bit
    _bAbort    : BOOL;                 // 中止撤离标记（eOpen 相区分出口）[-] | Abort evacuation flag
    _bCfgBad   : BOOL;                 // 组态非法当拍量 [-] | Illegal configuration
    _uInfo     : UDINT;                // 信息码每拍重算 | Info code per scan
    _uCycleCnt : UDINT;                // 循环计数锁存量 [次] | Cycle count latch
    rtStart    : R_TRIG;               // 启动沿实例，段 0 无条件刷新 | Start edge
    rtReset    : R_TRIG;               // 复位沿实例，段 0 无条件刷新 | Reset edge
    rtDone     : R_TRIG;               // 完成相沿实例（单拍化），段 0 无条件刷新 | Done phase edge for one-shot
    tonClampLp : TON;                  // 低压护模计时，段 0 无条件刷新 | LP protect timer
    tonClampHp : TON;                  // 高压锁模计时，段 0 无条件刷新 | HP clamp timer
    tonForce   : TON;                  // 锁模力闸等待计时，段 0 无条件刷新 | Force gate wait timer
    tonInject  : TON;                  // 射胶计时，段 0 无条件刷新 | Injection timer
    tonHold    : TON;                  // 保压计时，段 0 无条件刷新 | Hold timer
    tonCool    : TON;                  // 冷却计时，段 0 无条件刷新 | Cooling timer
    tonOpen    : TON;                  // 开模计时，段 0 无条件刷新 | Open timer
END_VAR
VAR CONSTANT
    DL_ICS_CNT_MAX : UDINT := 16#FFFF_FFFE;   // 计数饱和上限（留加 1 裕度）[次] | Count saturation limit
END_VAR

(* —— 段 0：当拍量派生 + 定时器与沿实例无条件周期刷新（R7 红线） —— *)
_bCfgBad := (tClampLpTimeout <= T#0S) OR (tClampHpTimeout <= T#0S) OR (tForceGateWait <= T#0S)
         OR (tInjectTimeout <= T#0S) OR (tHoldTime <= T#0S) OR (tCoolTime <= T#0S)
         OR (tOpenTimeout <= T#0S) OR (fClampForceMin <= 0.0) OR (fInjPressSp <= 0.0);  // 组态域闸 / Configuration gate
rtStart(CLK := bStartCmd);                                          // 启动沿每拍必调 / Start edge every scan
rtReset(CLK := bReset);                                             // 复位沿每拍必调 / Reset edge every scan
rtDone(CLK := (_eState = E_DL_IcsPhase.eDone));                     // 完成相沿每拍必调（单拍化） / Done edge every scan
tonClampLp(IN := (_eState = E_DL_IcsPhase.eClampLp), PT := tClampLpTimeout);   // 护模计时 / LP protect timing
tonClampHp(IN := (_eState = E_DL_IcsPhase.eClampHp), PT := tClampHpTimeout);   // 锁模计时 / HP clamp timing
tonForce(IN := (_eState = E_DL_IcsPhase.eClampHp) AND bMoldClosedLim AND (fClampForceAct < fClampForceMin), PT := tForceGateWait); // 力闸等待 / Force gate wait timing
tonInject(IN := (_eState = E_DL_IcsPhase.eInject), PT := tInjectTimeout);      // 射胶计时 / Injection timing
tonHold(IN := (_eState = E_DL_IcsPhase.eHold), PT := tHoldTime);               // 保压计时 / Hold timing
tonCool(IN := (_eState = E_DL_IcsPhase.eCool), PT := tCoolTime);               // 冷却计时 / Cooling timing
tonOpen(IN := (_eState = E_DL_IcsPhase.eOpen), PT := tOpenTimeout);            // 开模计时 / Open timing

(* —— 段 1：单拍量预清零（锁存量不入清单） —— *)
_uInfo := 16#0000_0000;                                             // 信息码每拍重算 / Info recomputed per scan
bCycleDone := rtDone.Q;                                             // 完成单拍出口（R_TRIG 单拍化） / Done one-shot outlet

(* —— 段 2：复位沿 + 组态域闸 —— *)
IF rtReset.Q AND (NOT _bCfgBad) THEN                                // 复位沿且组态合法 / Reset with legal config
    _bFault := FALSE;                                               // 清故障锁存位 / Clear fault latch
    _eCause := E_DL_IcsCause.eNone;                                 // 清成因 / Clear cause
    IF _eState = E_DL_IcsPhase.eFault THEN
        _eState := E_DL_IcsPhase.eIdle;                             // 故障相迁出唯一路径 / Sole fault exit
    END_IF
END_IF
IF _bCfgBad THEN                                                    // 组态域闸 / Configuration gate
    _bFault := TRUE;                                                // 置故障锁存 / Latch fault
    _eCause := E_DL_IcsCause.eCfgIllegal;                           // 归因组态 / Cause: config
END_IF

(* —— 段 3：中止优先拦截（安全撤离不置故障） —— *)
IF (NOT _bFault) AND bCycleAbort
   AND ((_eState = E_DL_IcsPhase.eClampLp) OR (_eState = E_DL_IcsPhase.eClampHp)
     OR (_eState = E_DL_IcsPhase.eInject)  OR (_eState = E_DL_IcsPhase.eHold)
     OR (_eState = E_DL_IcsPhase.eCool)) THEN
    _bAbort := TRUE;                                                // 中止标记置位（eOpen 出口区分） / Abort flag set
    _eState := E_DL_IcsPhase.eOpen;                                 // 直接进入开模安全撤离 / Enter open for safe evacuation
END_IF

(* —— 段 4：相位机（ENUM + CASE，ELSE 兜底） —— *)
CASE _eState OF

E_DL_IcsPhase.eIdle:
    IF rtStart.Q AND bMoldOpenLim AND (NOT _bFault) THEN
        _bAbort := FALSE;                                           // 新循环清中止标记 / Clear abort flag for new cycle
        _eState := E_DL_IcsPhase.eClampLp;                          // 开到位才允许启动 / Start only from fully open
    END_IF

E_DL_IcsPhase.eClampLp:
    IF _bFault THEN
        _eState := E_DL_IcsPhase.eFault;                            // 故障即时迁出 / Leave on fault
    ELSIF bMoldClosedLim THEN
        _eState := E_DL_IcsPhase.eClampHp;                          // 护模段合到位转高压 / Closed, switch to HP clamp
    ELSIF tonClampLp.Q THEN
        _bFault := TRUE;                                            // 护模超时出口（模具障碍） / LP protect timeout exit
        _eCause := E_DL_IcsCause.eClampLpTimeout;
        _eState := E_DL_IcsPhase.eFault;
    END_IF

E_DL_IcsPhase.eClampHp:
    IF _bFault THEN
        _eState := E_DL_IcsPhase.eFault;                            // 故障即时迁出 / Leave on fault
    ELSIF bMoldClosedLim AND (fClampForceAct >= fClampForceMin) THEN
        _eState := E_DL_IcsPhase.eInject;                           // 锁模力段间闸放行（边界①）/ Force gate passes, inject allowed
    ELSIF tonClampHp.Q AND (NOT bMoldClosedLim) THEN
        _bFault := TRUE;                                            // 锁模超时（未合到位） / HP clamp timeout, not closed
        _eCause := E_DL_IcsCause.eClampHpTimeout;
        _eState := E_DL_IcsPhase.eFault;
    ELSIF tonForce.Q THEN
        _bFault := TRUE;                                            // 力闸等待超时（含 NaN 挂窗路径，边界②）/ Force gate wait timeout
        _eCause := E_DL_IcsCause.eForceGateTimeout;
        _eState := E_DL_IcsPhase.eFault;
    END_IF

E_DL_IcsPhase.eInject:
    IF _bFault THEN
        _eState := E_DL_IcsPhase.eFault;                            // 故障即时迁出 / Leave on fault
    ELSIF fInjPressAct >= fInjPressSp THEN
        _eState := E_DL_IcsPhase.eHold;                             // 压力到切换点转保压 / Pressure at switchover, hold
    ELSIF tonInject.Q THEN
        _bFault := TRUE;                                            // 射胶超时（含熔胶未到位等待） / Injection timeout
        _eCause := E_DL_IcsCause.eInjectTimeout;
        _eState := E_DL_IcsPhase.eFault;
    END_IF

E_DL_IcsPhase.eHold:
    IF _bFault THEN
        _eState := E_DL_IcsPhase.eFault;                            // 故障即时迁出 / Leave on fault
    ELSIF tonHold.Q THEN
        _eState := E_DL_IcsPhase.eCool;                             // 保压时间到转冷却 / Hold elapsed, cool
    END_IF

E_DL_IcsPhase.eCool:
    IF _bFault THEN
        _eState := E_DL_IcsPhase.eFault;                            // 故障即时迁出 / Leave on fault
    ELSIF tonCool.Q THEN
        _eState := E_DL_IcsPhase.eOpen;                             // 冷却时间到开模 / Cool elapsed, open
    END_IF

E_DL_IcsPhase.eOpen:
    IF bMoldOpenLim THEN
        IF _bAbort THEN
            _uInfo := 16#0005_04DB;                                 // 信息级：中止撤离完成 / Info: abort evacuation done
            _bAbort := FALSE;                                       // 清中止标记 / Clear abort flag
            _eState := E_DL_IcsPhase.eIdle;                         // 撤离完成回待机（不计数） / Evacuated, no count
        ELSE
            _eState := E_DL_IcsPhase.eDone;                         // 正常开到位进完成相 / Normal open done
        END_IF
    ELSIF tonOpen.Q THEN
        _bFault := TRUE;                                            // 开模超时 / Open timeout
        _eCause := E_DL_IcsCause.eOpenTimeout;
        _eState := E_DL_IcsPhase.eFault;
    END_IF

E_DL_IcsPhase.eDone:
    IF _uCycleCnt < DL_ICS_CNT_MAX THEN
        _uCycleCnt := _uCycleCnt + 1;                               // 完成计数递增（本相仅驻留一拍） / Count increment, one-scan phase
    END_IF
    _uInfo := 16#0005_04DA;                                         // 信息级：循环完成台账 / Info: cycle done ledger
    _eState := E_DL_IcsPhase.eIdle;                                 // 完成即回待机（bCycleDone 由 rtDone 单拍化） / Back to idle, one-shot via rtDone

E_DL_IcsPhase.eFault:
    ;                                                               // 仅段 2 复位沿可迁出 / Only reset edge leaves

ELSE
    _bFault := TRUE;                                                // 非法相位兜底（R6）/ Illegal phase fallback
    _eCause := E_DL_IcsCause.eCfgIllegal;                           // 归因归并组态 / Cause folded to config
    _eState := E_DL_IcsPhase.eFault;

END_CASE

(* —— 段 5：故障锁存相位迁移闸 —— *)
IF _bFault AND (_eState <> E_DL_IcsPhase.eFault) THEN
    _eState := E_DL_IcsPhase.eFault;                                // 锁存即入故障相 / Latch enters fault phase
END_IF

(* —— 段 6：出口单点映射（名实同源；锁存码回放） —— *)
bClampFwd  := (_eState = E_DL_IcsPhase.eClampLp) OR (_eState = E_DL_IcsPhase.eClampHp);  // 合模输出两段 / Clamp output both segments
bClampHigh := (_eState = E_DL_IcsPhase.eClampHp);               // 高压输出 / HP output
bInjectOut := (_eState = E_DL_IcsPhase.eInject);                // 射胶输出 / Injection output
bHoldOut   := (_eState = E_DL_IcsPhase.eHold);                  // 保压输出 / Hold output
bCoolOut   := (_eState = E_DL_IcsPhase.eCool);                  // 冷却输出 / Cooling output
bOpenOut   := (_eState = E_DL_IcsPhase.eOpen);                  // 开模输出 / Open output
uCycleCnt  := _uCycleCnt;                                       // 计数镜像（锁存回放） / Count mirror
eState     := _eState;                                          // 相位出口 / Phase outlet
eCause     := _eCause;                                          // 成因出口 / Cause outlet
bError     := _bFault;                                          // 故障标志同源 / Error flag from latch
IF _bFault THEN
    nErrId := 16#0005_03B7;                                     // 故障锁存码回放 / Replay latched fault code
ELSE
    nErrId := _uInfo;                                           // 信息码 / Info code
END_IF

END_FUNCTION_BLOCK
